(* IEC 61131-3 sources: volt/packages/volt-lsp-iec/test-corpus/awa-palletizer/Device/Plc Logic/Application/Library Manager/L_MC1P_MotionControlBasic, 701 files *)

(* ---- L_MC1P_ABC_STATE.dut ---- *)
TYPE L_MC1P_ABC_STATE :
(
	STANDBY := 0,
	STOP := 1,
	HOMING := 2,
	JOGGING := 3,
	MOVEVEL := 4,
	MOVEABS := 5,
	MOVEREL := 6,
	EXTERNAL := 7,
	ERROR := 8,
	FINISHPOSITIONING := 9
);
END_TYPE

(* ---- L_MC1P_ABORTTRIGGERINPUT.dut ---- *)
TYPE L_MC1P_ABORTTRIGGERINPUT :
STRUCT
	PTRIGGER_REF : POINTER TO MC_TRIGGER_REF;
	EXECUTE : BOOL;
	PAUSEACTIVETP : BOOL;
END_STRUCT
END_TYPE

(* ---- L_MC1P_ABORTTRIGGEROUTPUT.dut ---- *)
TYPE L_MC1P_ABORTTRIGGEROUTPUT :
STRUCT
	DONE : BOOL;
	BUSY : BOOL;
	ERROR : BOOL;
	ERRORID : L_IE1P_Error;
END_STRUCT
END_TYPE

(* ---- L_MC1P_ADDITIONALCONFIGINFO.dut ---- *)
TYPE L_MC1P_ADDITIONALCONFIGINFO :
STRUCT
	LWIDENTDRIVESWITCHOFF : LWORD := 0;
	DWREVISION : DWORD := 0;
	DWMOTORRATEDSPEED : DWORD := 3000;
	LRREFCURRENTMOTOR : LREAL := 0;
	LRREFTORQUEMOTOR : LREAL := 1;
	LRMOTORRATEDTORQUE : LREAL := 1;
	LRTORQUELIMITFACTOR : LREAL := 1;
	LRINERTIAMOTOR : LREAL := 0.01;
	DWMOTORREVOLUTION : DWORD := 1;
	DWENCODERCRC : DWORD := 0;
	XRESETRETAINENCERRORAFTERMAINSWITCH : BOOL;
	XFEEDBACKABSPOSAVAILABLE : BOOL := TRUE;
	XVFCMODE : BOOL := FALSE;
	XTACIA402ADVANCED : BOOL := FALSE;
	WMCTRLMODEDRIVE : USINT := 1;
	XDRIVELOADENCODER : BOOL := FALSE;
	DWDRIVELOADENCODERFEEDBACKCONFIG : DWORD := 0;
	DWDRIVELOADENCODERORIENTATION : DWORD := 0;
	DWDRIVELOADENCODERCRC : DWORD := 0;
	XDEVICETRANSMITTIMESVALID : BOOL;
	LRDEVICETRANSMITTIMEACTPOSMS : LREAL;
	LRDEVICETRANSMITTIMESETPOSMS : LREAL;
END_STRUCT
END_TYPE

(* ---- L_MC1P_ADDITIONALLIMITS.dut ---- *)
TYPE L_MC1P_ADDITIONALLIMITS :
(
	NOTACTIVE := 0,
	ADDITIONALPOSLIMITS := 1
);
END_TYPE

(* ---- L_MC1P_AUTOTUNINGPARA.dut ---- *)
TYPE L_MC1P_AUTOTUNINGPARA :
STRUCT
	MAXVELOCITY : LREAL;
	MAXACCELERATION : LREAL := 0;
	MAXDISTANCE : LREAL := 0;
	MOVEMENTDISTANCE : LREAL := 0;
	STATE : WORD := 0;
	COMMANDIN : USINT;
	VPNFACTOR : WORD;
	TNNFACTOR : WORD;
	VPPFACTOR : WORD;
	VPPFACTOREXT : WORD;
	WAITINGTIME : LREAL;
END_STRUCT
END_TYPE

(* ---- L_MC1P_AVERAGEFILTERSETVALUESINPUT.dut ---- *)
TYPE L_MC1P_AVERAGEFILTERSETVALUESINPUT :
STRUCT
	WFILTERDEPTH : WORD;
	XMANIPULATETORQUE : BOOL := FALSE;
END_STRUCT
END_TYPE

(* ---- L_MC1P_AVERAGEFILTERSETVALUESOUTPUT.dut ---- *)
TYPE L_MC1P_AVERAGEFILTERSETVALUESOUTPUT :
STRUCT
	XINEQOUT : BOOL;
END_STRUCT
END_TYPE

(* ---- L_MC1P_AXIS_STATE.dut ---- *)
TYPE L_MC1P_AXIS_STATE :
(
	ERRORSTOP := 1,
	DISABLED := 2,
	STANDSTILL := 3,
	STOPPING := 4,
	DISCMOTION := 5,
	SYNCMOTION := 6,
	CONTMOTION := 7,
	HOMING := 8,
	SERVICE := 10
);
END_TYPE

(* ---- L_MC1P_AXISBASICCONTROLINPUT_INTERNAL.dut ---- *)
TYPE L_MC1P_AXISBASICCONTROLINPUT_INTERNAL :
STRUCT
	PAXIS : POINTER TO AXIS_REF;
	DISABLEMOVEFUNEXEC : BOOL;
	XDISABLEPOWERCALL : BOOL;
	XREGULATORON : BOOL;
	XRESETERROR : BOOL;
	XENABLEPOSITIVE : BOOL := TRUE;
	XENABLENEGATIVE : BOOL := TRUE;
	XDISABLESWLIMIT : BOOL;
	LROVERRIDE : LREAL := 1.0;
	LROVERRIDEACC : LREAL := 1.0;
	LROVERRIDEJERK : LREAL := 1.0;
	XSTOP : BOOL;
	LRSTOPDEC : LREAL;
	LRSTOPJERK : LREAL;
	XJOGGINGPOS : BOOL;
	XJOGGINGNEG : BOOL;
	LRJOGGINGSETVEL : LREAL := 3600;
	LRJOGGINGSETACC : LREAL := 36000;
	LRJOGGINGSETDEC : LREAL := 36000;
	LRJOGGINGSETJERK : LREAL := 0;
	LRJOGGINGSETJERKDEC : LREAL := 0;
	XCONTINUOUSUPDATE : BOOL;
	XFINISHPOSITIONING : BOOL;
	XQSPAPPLICATION : BOOL;
	XHALT : BOOL;
	XABORT : BOOL;
	XMOVEVELEXECUTE : BOOL;
	XMOVEABSEXECUTE : BOOL;
	XMOVERELEXECUTE : BOOL;
	LRSETPOS_DIST : LREAL;
	LRSETVEL : LREAL := 3600;
	LRSETACC : LREAL := 36000;
	LRSETDEC : LREAL := 36000;
	LRSETJERK : LREAL := 0;
	LRSETJERKDEC : LREAL := 0;
	ESETDIRECTION : MC_DIRECTION := MC_DIRECTION.mcPositiveDirection;
	XHOMEEXECUTE : BOOL;
	LRHOMEPOSITION : LREAL;
	XUSEHOMEEXTPARAMETER : BOOL;
	SCHOMEEXTPARAMETER : L_MC1P_HomeParameter;
	SCHOMEEXTTP : MC_TRIGGER_REF;
	XHOMEABSSWITCH : BOOL;
	XRESETHOMEPOSITION : BOOL;
	XMOVEVELENABLEOFFSETVEL : BOOL;
	LRMOVEVELOFFSETVEL : LREAL;
	XUSEABORTBEHAVIOURFORTM : BOOL;
	LRABORTDEC : LREAL;
	LRABORTJERK : LREAL;
END_STRUCT
END_TYPE

(* ---- L_MC1P_AXISBASICCONTROLINSTANCEDATA.dut ---- *)
TYPE L_MC1P_AXISBASICCONTROLINSTANCEDATA :
STRUCT
	XERROR : BOOL;
	EERRORID : L_IE1P_Error;
	XFUNBUSY : BOOL;
	XFUNDONE : BOOL;
	XFUNCOMMANDABORTED : BOOL;
	EFUNSTATEACT : L_MC1P_ABC_State;
	ABCFUNID : WORD;
	WPOWID : WORD;
	XEXIT : BOOL;
	XMOVEVELEXECUTEOLD : BOOL;
	XMOVEABSEXECUTEOLD : BOOL;
	XMOVERELEXECUTEOLD : BOOL;
	XFINISHPOSITIONINGOLD : BOOL;
	XHOMEEXECUTEOLD : BOOL;
	XJOGGINGNEGOLD : BOOL;
	XJOGGINGPOSOLD : BOOL;
	XSTOPOLD : BOOL;
	XHALTOLD : BOOL;
	XABORTOLD : BOOL;
	XPOWERROROLD : BOOL;
	XDISABLESWLIMITOLD : BOOL;
	XFUNDONEOLD : BOOL;
	XRESETHOMEPOSITIONOLD : BOOL;
	XSAVEMOVEVELDONE : BOOL;
	XACYCLICAXIS : BOOL;
	XQSPAPPLDETECTED : BOOL;
	FBSTOP_EXECUTE : BOOL;
	FBHALT_EXECUTE : BOOL;
	FBABORT_EXECUTE : BOOL;
	FBMOVEABS_EXECUTE : BOOL;
	FBMOVEVEL_EXECUTE : BOOL;
	FBMOVEREL_EXECUTE : BOOL;
	FBFINISHPOSITIONING_XFINISHPOSITIONING : BOOL;
	FBFINISHPOSITIONING_XENABLE : BOOL;
	FBJOG_XJOGPOSITIVE : BOOL;
	FBJOG_XJOGNEGATIVE : BOOL;
	FBHOME_EXECUTE : BOOL;
	FBSTOP_XINUSE : BOOL;
	FBHALT_XINUSE : BOOL;
	FBABORT_XINUSE : BOOL;
	FBMOVEABS_XINUSE : BOOL;
	FBMOVEVEL_XINUSE : BOOL;
	FBMOVEREL_XINUSE : BOOL;
	FBFINISHPOSITIONING_XINUSE : BOOL;
	FBJOG_XINUSE : BOOL;
	FBHOME_XINUSE : BOOL;
	XDRIVEENABLEDOLD_READMOTIONSTATE : BOOL;
	LRACTVELOCITYOLD_READMOTIONSTATE : LREAL;
	LRSETVELOCITYOLD_READMOTIONSTATE : LREAL;
	FBBASEOLD : POINTER TO L_MC1P_Template_ForAxis;
	FBSTOP_FBBASESTATUS : L_MC1P_Template_ForAxis;
	FBHALT_FBBASESTATUS : L_MC1P_Template_ForAxis;
	FBABORT_FBBASESTATUS : L_MC1P_Template_ForAxis;
	FBHOME_FBBASESTATUS : L_MC1P_Template_ForAxis;
	FBJOG_FBBASESTATUS : L_MC1P_Template_ForAxis;
	FBMOVEABS_FBBASESTATUS : L_MC1P_Template_ForAxis;
	FBMOVEVEL_FBBASESTATUS : L_MC1P_Template_ForAxis;
	FBMOVEREL_FBBASESTATUS : L_MC1P_Template_ForAxis;
	FBFINISHPOSITIONING_FBBASESTATUS : L_MC1P_Template_ForAxis;
	FBSETFASTSTOP_FBBASESTATUS : L_MC1P_Template_ForAxis;
	FBSETFASTSTOPINPUT : L_MC1P_SetQuickStopApplInput;
	FBSETFASTSTOP : L_MC1P_SetFastStop_Internal;
	FBSETFASTSTOPOUTPUT : L_MC1P_SetQuickStopApplOutput;
	FBRESET_FBBASESTATUS : L_MC1P_Template_ForAxis;
	FBRESET : L_MC1P_Reset_Internal;
	RESETINPUT : L_MC1P_ResetInput;
	RESETOUTPUT : L_MC1P_ResetOutput;
	FBSETOVERRIDE_FBBASESTATUS : L_MC1P_Template_ForAxis;
	FBSETOVERRIDE : L_MC1P_SetOverride_Internal;
	FBREADMOTIONSTATEINPUT : L_MC1P_ReadMotionStateInput;
	FBREADMOTIONSTATE_FBBASESTATUS : L_MC1P_Template_ForAxis;
	FBREADMOTIONSTATE : L_MC1P_ReadMotionState_Internal;
	FBREADMOTIONSTATEOUTPUT : L_MC1P_ReadMotionStateOutput;
	FBREADAXISERROR_FBBASESTATUS : L_MC1P_Template_ForAxis;
	FBREADAXISERROR : L_MC1P_ReadAxisError_Internal;
	FBREADAXISERRORINPUT : L_MC1P_ReadAxisErrorInput;
	FBREADAXISERROROUTPUT : L_MC1P_ReadAxisErrorOutput;
END_STRUCT
END_TYPE

(* ---- L_MC1P_AXISBASICCONTROLOUTPUT_INTERNAL.dut ---- *)
TYPE L_MC1P_AXISBASICCONTROLOUTPUT_INTERNAL :
STRUCT
	ECONTROLMODE : L_MC1P_ControlMode;
	XISHOMED : BOOL;
	XHWLIMITSWITCHNEG : BOOL;
	XHWLIMITSWITCHPOS : BOOL;
	XSWLIMITENABLED : BOOL;
	XSWLIMITSWITCHNEG : BOOL;
	XSWLIMITSWITCHPOS : BOOL;
	EAXISTYPE : L_MC1P_DriveType;
	EAXISSTATE : L_MC1P_AXIS_STATE := L_MC1P_AXIS_STATE.Disabled;
	XAXISREADY : BOOL;
	XAXISENABLED : BOOL;
	XAXISWARNING : BOOL;
	XAXISERROR : BOOL;
	EAXISERRORID : L_IE1P_Error;
	XDRIVEWARNING : BOOL;
	XDRIVEERROR : BOOL;
	DWDRIVEERRORID : DWORD;
	LRACTPOS : LREAL;
	LRACTVEL : LREAL;
	LRSETPOSOUT : LREAL;
	LRSETVELOUT : LREAL;
	LRACTFOLLOWINGERROR : LREAL;
	XCONSTANTVELOCITY : BOOL;
	XACCELERATING : BOOL;
	XDECELERATING : BOOL;
	XDIRECTIONPOSITIVE : BOOL;
	XDIRECTIONNEGATIVE : BOOL;
	XINPOSITION : BOOL;
	XAXISAVAILABLE : BOOL;
	XSTANDSTILLSETVELOCITY : BOOL;
	XSTANDSTILLACTVELOCITY : BOOL;
	XAXISREADYTOSWITCHON : BOOL;
	XAXISREADYFORMOTION : BOOL;
	XERROR : BOOL;
	EERRORID : L_IE1P_Error;
	XFUNBUSY : BOOL;
	XFUNDONE : BOOL;
	XFUNCOMMANDABORTED : BOOL;
	EFUNSTATEACT : L_MC1P_ABC_State;
	XSTOACTIVE : BOOL;
END_STRUCT
END_TYPE

(* ---- L_MC1P_AXISEXTENSIONTYPES.dut ---- *)
TYPE L_MC1P_AXISEXTENSIONTYPES :
(
	EMPTY := 0,
	HL9400_ECAT := 1,
	HL9400_CAN := 2,
	I500_ECAT := 3,
	I500_CAN := 4,
	I700 := 5,
	I750 := 6,
	I950 := 7,
	I950ADV := 8,
	I950_DRIVE := 9,
	I950_DRIVECIA := 10,
	GENERICDRIVE := 11,
	ENCFREE := 101,
	ENCIO_BPB := 102,
	ENCIO_ECAT := 103,
	ENCI900_ECAT := 104,
	ENCI900_DRIVE := 105,
	ENCI900_DRIVECIA := 106,
	ENCI500_ECAT := 107
);
END_TYPE

(* ---- L_MC1P_AXISFUNCTION.dut ---- *)
TYPE L_MC1P_AXISFUNCTION :
(
	SIMPLEMODE := 1,
	PLI := 2,
	MOL := 3,
	POSCTRLADAPT := 4,
	SPEEDCTRLADAPT := 5,
	SPEEDCTRLLOAD := 6,
	BRAKEGRINDIN := 7,
	BRAKETEST := 8,
	BASICBRAKECTRLONLYINDRIVE := 9,
	FLEXIBLEMAPPING := 10,
	ZEROPULS2NDFEEDBACK := 11,
	FDBSTATUSBITSAVAILABLE := 12,
	AUTOTUNING := 13,
	PARSAVEINDRIVE := 14,
	WAITFORAXISDETECTION := 15
);
END_TYPE

(* ---- L_MC1P_AXISGUID.dut ---- *)
TYPE L_MC1P_AXISGUID :
STRUCT
	ADWDATA : ARRAY [1..4] OF DWORD;
END_STRUCT
END_TYPE

(* ---- L_MC1P_AXISINTERFACEINPUT.dut ---- *)
TYPE L_MC1P_AXISINTERFACEINPUT :
STRUCT
	XENABLE : BOOL;
	EXTCONTROLLER : L_MC1P_IControllerInterface;
END_STRUCT
END_TYPE

(* ---- L_MC1P_AXISINTERFACEOUTPUT.dut ---- *)
TYPE L_MC1P_AXISINTERFACEOUTPUT :
STRUCT
	XVALID : BOOL;
	XBUSY : BOOL;
	XERROR : BOOL;
	EERRORID : L_IE1P_Error;
END_STRUCT
END_TYPE

(* ---- L_MC1P_AXISPROPERTIES.dut ---- *)
TYPE L_MC1P_AXISPROPERTIES :
STRUCT
	XVIRTUAL : BOOL := FALSE;
	XTPSUPPORTED : BOOL := FALSE;
	XTPWITHTIMESTAMP : BOOL := FALSE;
	SNTPMAXCHANNEL : SINT := 0;
	XSUPPORTBRAKE : BOOL := FALSE;
	XSUPPORTDCBRAKE : BOOL := FALSE;
	XCHECKCOMMUNICATIONSTATE : BOOL := TRUE;
	XDRIVEHOMINGSUPPORTED : BOOL := FALSE;
	XTACIAADVANCED : BOOL := FALSE;
	BYDELAYLIMITDRIVEOPERATIONENABLED : BYTE := 2;
	LRTRANSMITCYCLESACTPOS : LREAL;
	LRTRANSMITCYCLESSETPOS : LREAL;
	DWTPDELAYACTPOS : DWORD;
	XFORWARDECATSLAVEERROR : BOOL := FALSE;
	XFORCEACYCLICMODE : BOOL := FALSE;
	WOFFSETDRIVEPARA : WORD := 0;
END_STRUCT
END_TYPE

(* ---- L_MC1P_AXISRETAININFO.dut ---- *)
TYPE L_MC1P_AXISRETAININFO :
STRUCT
	MEMTYPE : BYTE;
	MEMVERSION : BYTE;
	MEMLENGTH : WORD;
END_STRUCT
END_TYPE

(* ---- L_MC1P_AXISRETAININFORMATION.dut ---- *)
TYPE L_MC1P_AXISRETAININFORMATION :
STRUCT
	AXISGUID : L_MC1P_AxisGUID;
	ITFRETAIN : L_MC1P_IRetainFunction;
	PDATA : POINTER TO DWORD;
	PDATAMIRROR : POINTER TO DWORD;
END_STRUCT
END_TYPE

(* ---- L_MC1P_AXISSIMIODATA.dut ---- *)
TYPE L_MC1P_AXISSIMIODATA :
STRUCT
	XSTO : BOOL;
	XDIGIN1 : BOOL;
	XDIGIN2 : BOOL;
	XSTIMULATEERROR : BOOL;
	DWERRORCODE : DWORD;
	XQSPONERROR : BOOL;
	XSTIMULATEWARNING : BOOL;
	DWWARNINGCODE : DWORD;
	ETPMODE : UINT := 0;
	LRTPDISTANCE : LREAL;
	LRTPDISTANCEINTERNAL : LREAL;
	XSTIMULATEFEEDBACKCHANGED : BOOL;
END_STRUCT
END_TYPE

(* ---- L_MC1P_AXISSIMULATIONPDODATAFROMDRIVE.dut ---- *)
TYPE L_MC1P_AXISSIMULATIONPDODATAFROMDRIVE :
STRUCT
	UICIASTATUSWORD : UINT;
	UILENZESTATUSWORD : UINT;
	SIMODEOFOPERATIONDISP : SINT;
	UIERRORCODE : UINT;
	UITEXTREFID : UINT;
	DIVELACTVALUE : DINT;
	ITORQUEACTVALUE : INT;
	DIPOSACTVALUE : DINT;
	DIFOLLOWINGERRORACTVALUE : DINT;
	IVLACTUALVEL : INT;
	UITPSTATUS : UINT;
	DITPPOS1POSVALUE : DINT;
	DITPPOS1NEGVALUE : DINT;
	DITPPOS2POSVALUE : DINT;
	DITPPOS2NEGVALUE : DINT;
	UILENZESTATUSWORD2 : UINT;
	UDIDIGITALINPUTS : UDINT;
END_STRUCT
END_TYPE

(* ---- L_MC1P_AXISSIMULATIONPDODATAFROMDRIVESCALED.dut ---- *)
TYPE L_MC1P_AXISSIMULATIONPDODATAFROMDRIVESCALED :
STRUCT
	UICIASTATUSWORD : UINT;
	UILENZESTATUSWORD : UINT;
	SIMODEOFOPERATIONDISP : SINT;
	UIERRORCODE : UINT;
	UITEXTREFID : UINT;
	LRVELACTVALUE : LREAL;
	LRTORQUEACTVALUE : LREAL;
	LRPOSACTVALUE : LREAL;
	LRFOLLOWINGERRORACTVALUE : LREAL;
	UITPSTATUS : UINT;
	LRTPPOS1POSVALUE : LREAL;
	LRTPPOS1NEGVALUE : LREAL;
	LRTPPOS2POSVALUE : LREAL;
	LRTPPOS2NEGVALUE : LREAL;
	UILENZESTATUSWORD2 : UINT;
	UDIDIGITALINPUTS : UDINT;
END_STRUCT
END_TYPE

(* ---- L_MC1P_AXISSIMULATIONPDODATATODRIVE.dut ---- *)
TYPE L_MC1P_AXISSIMULATIONPDODATATODRIVE :
STRUCT
	UICTRLWORD : UINT;
	UILENZECTRLWORD : UINT;
	SIMODEOFOPERATION : SINT;
	ITORQUEOFFSET : INT;
	DITARGETPOSITION : DINT;
	DIVELOCITYOFFSET : DINT;
	ISPDCTRL_ILOADVALUE : INT;
	ITARGETTORQUE : INT;
	DITARGETVELOCITY : DINT;
	IVLTARGETVEL : INT;
	UITPFUNCTION1 : UINT;
	UIPOSTORQUELIMIT : UINT;
	UINEGTORQUELIMIT : UINT;
	DIUPPERSPEEDLIMIT : DINT;
	DILOWERSPEEDLIMIT : DINT;
END_STRUCT
END_TYPE

(* ---- L_MC1P_AXISSIMULATIONPDODATATODRIVESCALED.dut ---- *)
TYPE L_MC1P_AXISSIMULATIONPDODATATODRIVESCALED :
STRUCT
	UICTRLWORD : UINT;
	UILENZECTRLWORD : UINT;
	SIMODEOFOPERATION : SINT;
	LRSETPOSITION : LREAL;
	LRSETVELOCITY : LREAL;
	LRSETTORQUE : LREAL;
	LRSPDCTRL_ILOADVALUE : LREAL;
	LRVLTARGETVELOCITY : LREAL;
	UITPFUNCTION1 : UINT;
	LRPOSTORQUELIMIT : LREAL;
	LRNEGTORQUELIMIT : LREAL;
	LRUPPERSPEEDLIMIT : LREAL;
	LRLOWERSPEEDLIMIT : LREAL;
END_STRUCT
END_TYPE

(* ---- L_MC1P_AXISSIMULATIONSDODATA.dut ---- *)
TYPE L_MC1P_AXISSIMULATIONSDODATA :
STRUCT
	LRRATEDMOTORTORQUE : LREAL := 0.6;
	LRRATEDMOTORSPEED : LREAL := 4050;
	LRINERTIAMOTOR : LREAL := 0.14;
	LRINERTIALOAD : LREAL := 0;
	LRMOTORRATEDCURRENT : LREAL := 1.8;
	LRMAXMOTORSPEED : LREAL := 6075;
	BYMCTRLMODE : BYTE := 1;
	LRVP_SPEEDCTRL : LREAL := 0.00045;
	LRTN_SPEEDCTRL : LREAL := 12.8;
	LRVP_POSCTRL : LREAL := 28.4;
	LRPOSCTRLOUTPUTLIMITATION : LREAL := 480000;
	UIINSABILITYVALUE : UINT;
	UIINSABILITYINDICATOR : USINT;
	USISWITCHINGFREQUENCY : USINT := 1;
	LRPOSCTRLADAPT : LREAL := 100.0;
	LRSPEEDCTRLADAPT : LREAL := 100.0;
	LRMAXTORQUE : LREAL := 250.0;
	LRSPEEDFILTERTIME : LREAL := 0.3;
	WNBRORREVOLUTION : WORD := 1;
	DWINKPERREV : DWORD := 65536;
	DWENCODERCRC : DWORD := 1234;
	DWENCODERCRCLOAD : DWORD := 4567;
	USIBRAKEMODE : USINT := 2;
	UIBRAKESRCOFSTARTINGTORQUE : UINT := 1;
	LRBRAKEDETECTEDSTARTINGTORQUE : LREAL := 0;
	LRBRAKERELEASINGTIME : LREAL := 0.1;
	LRBRAKECLOSINGTIME : LREAL := 0.1;
	USIBRAKEOVERRIDE : USINT := 0;
	LRSTARTTORQUE : LREAL;
	UIBRAKELOGICSTATE : UINT;
	UICONTROLMODECIA402ADVANCED : UINT := 0;
	LRVP_LOADPOSCTRL : LREAL := 20.0;
	SIIPOTIMEEXP : SINT;
	USIIPOTIME : USINT;
	UIQSPOPTION : UINT;
	UDIPOSITIONREACHEDWINDOW : UDINT := 1000;
	UDIQSPDECELERATION : UDINT := 2147483647;
	DWREVISIONNBR : DWORD := 16#20000;
	DWFIRSTSYNCTIME : DWORD;
	USISPEEDERRORRESPONSE : USINT;
	SSWVERSION : STRING(50) := '1.7.5.2420 (release)';
	USIDISABLEPDOS : USINT;
	USIDRIVECOMMAND_0X2825 : USINT;
	UDIMAINSWITCHINGCYCLES_0X2D81_4 : UDINT := 666;
	USIPOSSETMODE_0X2984 : USINT;
	LRVLACCDELTASPEED : LREAL := 0;
	LRVLACCDELTATIME : LREAL := 10;
	LRVLDECDELTASPEED : LREAL := 0;
	LRVLDECDELTATIME : LREAL := 0;
	BYDISABLEDEVICE : BYTE;
	DIADDSPEEDLIMITATION : DINT := 0;
	AUIGAINCHARACTERISTIC : ARRAY [1..11] OF WORD := [10, 100, 100, 100, 1000, 100, 2000, 100, 5000, 100, 0];
END_STRUCT
END_TYPE

(* ---- L_MC1P_AXISSLOT.dut ---- *)
TYPE L_MC1P_AXISSLOT :
(
	AXISA := 16#0,
	AXISB := 16#800
);
END_TYPE

(* ---- L_MC1P_AXISTYPE.dut ---- *)
TYPE L_MC1P_AXISTYPE :
(
	UNKNOWN := 0,
	AXISREF := 1,
	AXISKINEMATIC := 2,
	AXISGROUP := 3
);
END_TYPE

(* ---- L_MC1P_BACKLASHCONTACTSTATE.dut ---- *)
TYPE L_MC1P_BACKLASHCONTACTSTATE :
(
	NOCONTACT := 0,
	NEGATIVECONTACT := 1,
	POSITIVECONTACT := 2
);
END_TYPE

(* ---- L_MC1P_BASICACTUATINGSPEEDINPUT.dut ---- *)
TYPE L_MC1P_BASICACTUATINGSPEEDINPUT :
STRUCT
	XENABLEINTERNALCONTROL : BOOL := FALSE;
	XREGULATORON : BOOL := FALSE;
	XRESETERROR : BOOL := FALSE;
	XSETDRIVEQSP : BOOL := FALSE;
	XENABLESETVEL : BOOL := FALSE;
	XINVERTDIRECTION : BOOL := FALSE;
	LRSETVEL : LREAL := 0.0;
	LRSETACC : LREAL := 0.0;
	LRSETDEC : LREAL := 0.0;
END_STRUCT
END_TYPE

(* ---- L_MC1P_BASICACTUATINGSPEEDOUTPUT.dut ---- *)
TYPE L_MC1P_BASICACTUATINGSPEEDOUTPUT :
STRUCT
	XINTERNALCONTROLACTIVE : BOOL;
	XBUSY : BOOL;
	XERROR : BOOL;
	EERRORID : L_IE1P_Error;
	XCOMMUNICATIONOK : BOOL;
	XAXISREADY : BOOL;
	XAXISENABLED : BOOL;
	XDRIVEWARNING : BOOL;
	XDRIVEERROR : BOOL;
	DWDRIVEERRORID : DWORD;
	XDRIVEQSPACTIVE : BOOL;
	LRACTVEL : LREAL;
	XDIRECTIONPOSITIVE : BOOL;
	XDIRECTIONNEGATIVE : BOOL;
	WDIGITALINPUTS : WORD;
END_STRUCT
END_TYPE

(* ---- L_MC1P_BRAKEAUTOSTATE.dut ---- *)
TYPE L_MC1P_BRAKEAUTOSTATE :
(
	AS_IDLE,
	AS_RAMPDOWN,
	AS_CLOSINGBRAKE,
	AS_INITBRAKECLOSE,
	AS_BRAKECLOSED,
	AS_RELEASINGBRAKE,
	AS_SUPERVISORMODE,
	AS_DIRECTCONTROL
);
END_TYPE

(* ---- L_MC1P_BRAKECMDBRAKEGRINDINPARA.dut ---- *)
TYPE L_MC1P_BRAKECMDBRAKEGRINDINPARA :
STRUCT
	MOTORSPEED : INT := 1000;
	RAMPTIME : INT := 1000;
	ONTIME : INT := 500;
	OFFTIME : INT := 500;
	CYCLES : WORD := 4;
	GRINDINCONTROL : BYTE;
	MODE : USINT;
	CYCLESOUT : WORD;
	STATE : WORD;
	POSLIMIT1 : LREAL;
	POSLIMIT2 : LREAL;
END_STRUCT
END_TYPE

(* ---- L_MC1P_BRAKECMDBRAKETESTPARA.dut ---- *)
TYPE L_MC1P_BRAKECMDBRAKETESTPARA :
STRUCT
	MOTORTORQUE : DINT := 0;
	RAMPTIME : INT := 1000;
	HOLDTIME : INT := 4000;
	POSTHRESHOLD : INT;
	STATE : WORD := 0;
	WBRAKETESTMODE : USINT;
END_STRUCT
END_TYPE

(* ---- L_MC1P_BRAKECTRL.dut ---- *)
TYPE L_MC1P_BRAKECTRL :
STRUCT
	XDISABLEPHIERR : BOOL;
	XBRAKEFQSP : BOOL;
	XTORQUETIMEOUT : BOOL;
	XRELEASED : BOOL;
	XOUTPUTRELEASEOLD : BOOL;
	XOBSERVE : BOOL;
	XMODULENOTOK : BOOL;
	XEXTSIGNOTOK : BOOL;
	XMODULEFEEDBACK : BOOL;
	XBRAKEOPENED : BOOL;
	XBRAKECLOSED : BOOL;
	XINVERTBRAKE : BOOL;
	XINVERTBRAKEOLD : BOOL;
	XUVDETECTEDOLD : BOOL;
	XACTSPEEDBELOWMINSPEED : BOOL;
	XBIT15 : BOOL;
END_STRUCT
END_TYPE

(* ---- L_MC1P_BRAKEERRORCODES.dut ---- *)
TYPE L_MC1P_BRAKEERRORCODES :
(
	EC_POSITIONDRIFT := 3,
	EC_POSITIONDRIFTCINH := 11,
	EC_RAMPWATCH := 4,
	EC_ERRORMODULE := 5,
	EC_ERROREXTSIGNAL := 13,
	EC_ERRORTORQUETIMEOUT := 18,
	EC_ERRORBRAKESTATEINVALID := 19,
	EC_ERRORBRAKEMODEINVALID := 20,
	EC_TORQUELIMITED := 30
);
END_TYPE

(* ---- L_MC1P_BRAKEGRINDININPUT.dut ---- *)
TYPE L_MC1P_BRAKEGRINDININPUT :
STRUCT
	XEXECUTE : BOOL;
	EMODE : L_MC1P_GrindInMode := L_MC1P_GrindInMode.CwCcw;
	EADDITIONALLIMITS : L_MC1P_AdditionalLimits := L_MC1P_AdditionalLimits.NotActive;
	LRPOSLIMIT1 : LREAL := 0;
	LRPOSLIMIT2 : LREAL := 0;
	LRMOTORSPEED : LREAL := 60.0;
	LRRAMPTIME : LREAL := 1.0;
	LRONTIME : LREAL := 0.5;
	LROFFTIME : LREAL := 0.5;
	WCYCLES : WORD := 4;
	XEXTERNALFAN : BOOL := FALSE;
	XFINISHINSTARTPOS : BOOL := FALSE;
	XUSEAXISPARAMETER : BOOL := FALSE;
	XDISABLEHOMEPOSCHECK : BOOL;
	XGRINDINVELOCITYMODE : BOOL;
	XCYCLESSETBYPARAMETER : BOOL;
	WCYCLESCW : WORD := 2;
	WCYCLESCCW : WORD := 2;
	XALLOWEXECUTIONFORKINEMATICSLAVE : BOOL;
	XABORT : BOOL;
END_STRUCT
END_TYPE

(* ---- L_MC1P_BRAKEGRINDINOUTPUT.dut ---- *)
TYPE L_MC1P_BRAKEGRINDINOUTPUT :
STRUCT
	XDONE : BOOL;
	XBUSY : BOOL;
	XACTIVE : BOOL;
	XCOMMANDABORTED : BOOL;
	XERROR : BOOL;
	EERRORID : L_IE1P_Error;
	WCYCLESOUT : WORD;
	ESTATE : L_MC1P_BrakeGrindInState := L_MC1P_BrakeGrindInState.NotActive;
	XGRINDINABORTEDINSTANDSTILL : BOOL;
END_STRUCT
END_TYPE

(* ---- L_MC1P_BRAKEGRINDINSTATE.dut ---- *)
TYPE L_MC1P_BRAKEGRINDINSTATE :
(
	NOTACTIVE := 0,
	INIT := 1,
	BRAKEGRINDIN := 3,
	DONE := 4,
	ERROR := 5,
	ABORTED := 6,
	BRAKEGRINDINFOLLOWER := 20
);
END_TYPE

(* ---- L_MC1P_BRAKEINTERFACEINPUT.dut ---- *)
TYPE L_MC1P_BRAKEINTERFACEINPUT :
STRUCT
	XENABLE : BOOL;
	XRELEASEBRAKE : BOOL;
	LRTORQUEADD : LREAL;
	XBRAKEMODEACTIVATE : BOOL;
	EBRAKEMODE : L_MC1P_BrakeMode;
END_STRUCT
END_TYPE

(* ---- L_MC1P_BRAKEINTERFACEOUTPUT.dut ---- *)
TYPE L_MC1P_BRAKEINTERFACEOUTPUT :
STRUCT
	XVALID : BOOL;
	XBUSY : BOOL;
	XERROR : BOOL;
	EERRORID : L_IE1P_Error;
	XBRAKERELEASEOUT : BOOL;
	XBRAKERELEASED : BOOL;
	LRACTTORQUE : LREAL;
	LRSTARTINGTORQUESAVED : LREAL;
	LRSTARTINGTORQUEEFFECTIVE : LREAL;
	EBRAKEMODEACTIVE : L_MC1P_BrakeMode;
END_STRUCT
END_TYPE

(* ---- L_MC1P_BRAKELOGICSTATE.dut ---- *)
TYPE L_MC1P_BRAKELOGICSTATE :
(
	OFF := 0,
	WAITON := 1,
	SELECTPRETORQUE := 10,
	LOADPRETORQUE := 11,
	OPENBRAKE := 20,
	OPERATION := 30,
	CLOSEBRAKE := 40,
	TURNOFF := 50
);
END_TYPE

(* ---- L_MC1P_BRAKEMODE.dut ---- *)
TYPE L_MC1P_BRAKEMODE :
(
	OFF := 0,
	MANUALCONTROL_PLC := 1,
	AUTOMATIC_PLC := 2
);
END_TYPE

(* ---- L_MC1P_BRAKEOUTSTATE.dut ---- *)
TYPE L_MC1P_BRAKEOUTSTATE :
STRUCT
	XBRAKECONTROLACTIVE : BOOL;
	XMODULEOPERATION : BOOL;
	XBRAKEOUTSTATE : BOOL;
	XTORQUECTRLACTIVE : BOOL;
	XBRAKECINH : BOOL;
	XERRORACTIVE : BOOL;
	XGRINDINACTIVE : BOOL;
	XTORQUETESTACTIVE : BOOL;
	XMANOPERATION : BOOL;
	XAUTOPERATION : BOOL;
	XERROREXTFEEDBACK : BOOL;
	XERRORPOSDRIFT : BOOL;
	XERRORBRAKEMODULE : BOOL;
	XINFOTIMEOUTACTIVATE : BOOL;
	XGRINDINDONE : BOOL;
	XTORQUETESTDONE : BOOL;
	XERRORTORQUECTRL : BOOL;
	XACTSPEEDBELOWMIN : BOOL;
	XERRORTORQUELIMITED : BOOL;
END_STRUCT
END_TYPE

(* ---- L_MC1P_BRAKEPARA.dut ---- *)
TYPE L_MC1P_BRAKEPARA :
STRUCT
	LRRELEASETIME : LREAL;
	LRACTIVATIONTIME : LREAL;
	DWBRAKEMODE : DWORD;
	ESELBRAKEMODE : DWORD;
	LRSAMPLEDBRAKETORQUE : LREAL;
	LREFFECTIVESTARTINGTORQUE : LREAL;
	ALRMSTARTVALUE : ARRAY [1..2] OF LREAL;
	LRBRAKERAMPTIME : LREAL;
	XBRAKEACCDEPENDING : BOOL;
	WSOURCESTARTVALUE : WORD;
END_STRUCT
END_TYPE

(* ---- L_MC1P_BRAKESTATE.dut ---- *)
TYPE L_MC1P_BRAKESTATE :
(
	EBS_DEFAULT := 0,
	EBS_BRAKECLOSED,
	EBS_BRAKEOPEN,
	EBS_BRAKESWITCHING,
	EBS_BRAKEOBSERVATION,
	EBS_BRAKEAUTO,
	EBS_BRAKEAUTOGSB,
	EBS_BRAKEAUTOSUPERVISOR,
	EBS_BRAKEMANUAL,
	EBS_BRAKEOFF,
	EBS_STATESWITCH,
	EBS_STATEOPERATION
);
END_TYPE

(* ---- L_MC1P_BRAKETESTINPUT.dut ---- *)
TYPE L_MC1P_BRAKETESTINPUT :
STRUCT
	XEXECUTE : BOOL;
	LRMOTORTORQUE : LREAL := 0;
	LRRAMPTIME : LREAL := 1.0;
	LRHOLDTIME : LREAL := 4.0;
	LRPOSTHRESHOLD : LREAL;
	EDIRECTION : MC_DIRECTION := MC_DIRECTION.mcCurrentDirection;
	EMODE : L_MC1P_BrakeTestMode := L_MC1P_BrakeTestMode.NoLoadTorque;
	XUSEAXISPARAMETER : BOOL := FALSE;
	XABORT : BOOL;
	XALLOWEXECUTIONFORKINEMATICSLAVE : BOOL;
END_STRUCT
END_TYPE

(* ---- L_MC1P_BRAKETESTMODE.dut ---- *)
TYPE L_MC1P_BRAKETESTMODE :
(
	NOLOADTORQUE := 0,
	LOADTORQUEIDENTIFICATION := 1
);
END_TYPE

(* ---- L_MC1P_BRAKETESTOUTPUT.dut ---- *)
TYPE L_MC1P_BRAKETESTOUTPUT :
STRUCT
	XDONE : BOOL;
	XBUSY : BOOL;
	XACTIVE : BOOL;
	XCOMMANDABORTED : BOOL;
	XERROR : BOOL;
	EERRORID : L_IE1P_Error;
	LRIDENTIFIEDTORQUE : LREAL;
	LRACTPOSTHRESHOLD : LREAL;
	LRACTMOTORTORQUE : LREAL;
	ESTATE : L_MC1P_BrakeTestState := L_MC1P_BrakeTestState.NotActive;
END_STRUCT
END_TYPE

(* ---- L_MC1P_BRAKETESTSTATE.dut ---- *)
TYPE L_MC1P_BRAKETESTSTATE :
(
	NOTACTIVE := 0,
	INIT := 1,
	TORQUEIDENTIFICATION := 2,
	BRAKETEST := 3,
	DONE := 4,
	ERROR := 5,
	ABORTED := 6,
	BRAKETESTFOLLOWER := 20
);
END_TYPE

(* ---- L_MC1P_BUFFERDATA.dut ---- *)
TYPE L_MC1P_BUFFERDATA :
STRUCT
	LRBUFFERPOSITIONPOS : LREAL;
	LRBUFFERPOSITIONNEG : LREAL;
	LRBUFFERVELPOS : LREAL;
	LRBUFFERVELNEG : LREAL;
END_STRUCT
END_TYPE

(* ---- L_MC1P_CHANGEMACHINEDATAINPUT.dut ---- *)
TYPE L_MC1P_CHANGEMACHINEDATAINPUT :
STRUCT
	XEXECUTE : BOOL;
	XSETFEEDCONSTANT : BOOL;
	LRFEEDCONSTANT : LREAL := 360.0;
	XSETGEARFACTOR : BOOL;
	DWGEARDENOMINATOR : DWORD := 1;
	DWGEARNUMERATOR : DWORD := 1;
	XSETADDGEARFACTOR : BOOL;
	DWADDGEARDENOMINATOR : DWORD := 1;
	DWADDGEARNUMERATOR : DWORD := 1;
	XSETPOSRESOLUTION : BOOL;
	DWPOSRESOLUTION : DWORD := 65536;
	XSETORIENTATION : BOOL;
	XORIENTATION : BOOL := FALSE;
	XSETTRAVERSINGRANGE : BOOL;
	ETRAVERSINGRANGE : L_MC1P_TraversingRange := L_MC1P_TraversingRange.Limited;
	XSETCYCLELENGTH : BOOL;
	LRCYCLELENGTH : LREAL := 360.0;
END_STRUCT
END_TYPE

(* ---- L_MC1P_CHANGEMACHINEDATAOUTPUT.dut ---- *)
TYPE L_MC1P_CHANGEMACHINEDATAOUTPUT :
STRUCT
	XDONE : BOOL;
	XBUSY : BOOL;
	XERROR : BOOL;
	EERRORID : L_IE1P_Error;
END_STRUCT
END_TYPE

(* ---- L_MC1P_CINHHANDLINGINPUT.dut ---- *)
TYPE L_MC1P_CINHHANDLINGINPUT :
STRUCT
	XENABLE : BOOL;
	XSTAYINLASTSTATE : BOOL;
	XMOVELASTSETPOS : BOOL;
	LRWINDOWPOS : LREAL;
	LRWINDOWNEG : LREAL;
	LRSETVEL : LREAL;
	LRSETACC : LREAL;
	LRSETDEC : LREAL;
	LRSETJERK : LREAL;
	EDIRECTION : MC_DIRECTION;
END_STRUCT
END_TYPE

(* ---- L_MC1P_CINHHANDLINGOUTPUT.dut ---- *)
TYPE L_MC1P_CINHHANDLINGOUTPUT :
STRUCT
	XDONE : BOOL;
	XBUSY : BOOL;
	XACTIVE : BOOL;
	XERROR : BOOL;
	EERRORID : L_IE1P_Error;
	XREADYTOCONTINUE : BOOL;
	XINSIDEPOSWINDOW : BOOL;
	XINSIDEACTPOSWINDOW : BOOL;
	EAXISSTATEREAL : L_MC1P_AXIS_STATE := L_MC1P_AXIS_STATE.Disabled;
	LRDISTANCE : LREAL;
END_STRUCT
END_TYPE

(* ---- L_MC1P_CLASSID.dut ---- *)
TYPE L_MC1P_CLASSID :
(
	AXIS_REF := (L_MC1P_Internal.cdiEnumStartValue + 2),
	AXISBASICCONTROLV2 := (L_MC1P_Internal.cdiEnumStartValue + 3)
);
END_TYPE

(* ---- L_MC1P_COMPENSATIONMODE.dut ---- *)
TYPE L_MC1P_COMPENSATIONMODE :
(
	OFF := 0,
	AUTOMATICSET := 1,
	AUTOMATICACT := 2,
	MANUALLY := 3
);
END_TYPE

(* ---- L_MC1P_CONTROLAXIS.dut ---- *)
TYPE L_MC1P_CONTROLAXIS :
STRUCT
	XENABLEOPERATION : BOOL;
	XRESETERROR : BOOL;
	XQSPAPPLICATION : BOOL;
	XJOGPOS : BOOL;
	XJOGNEG : BOOL;
	LRJOGOVERRIDE : LREAL := 1.0;
	LRJOGDISTANCE : LREAL := 10;
	XRESETHOMEPOSITION : BOOL;
END_STRUCT
END_TYPE

(* ---- L_MC1P_CONTROLMODE.dut ---- *)
TYPE L_MC1P_CONTROLMODE :
(
	POSCTRLDRIVE := 0,
	POSCTRLPLC := 1,
	SPEEDCTRLDRIVE := 10,
	TORQUECTRLDRIVE := 20
);
END_TYPE

(* ---- L_MC1P_CONTROLMODESET.dut ---- *)
TYPE L_MC1P_CONTROLMODESET :
(
	POSCTRLDRIVE := 0,
	POSCTRLPLC := 1,
	SPEEDCTRLDRIVE := 10
);
END_TYPE

(* ---- L_MC1P_CTRLABC.dut ---- *)
TYPE L_MC1P_CTRLABC :
STRUCT
	XREGULATORON : BOOL;
	XRESETERROR : BOOL;
	XENABLEPOSITIVE : BOOL := TRUE;
	XENABLENEGATIVE : BOOL := TRUE;
	XDISABLESWLIMIT : BOOL;
	LROVERRIDE : LREAL := 1.0;
	LROVERRIDEACC : LREAL := 1.0;
	LROVERRIDEJERK : LREAL := 1.0;
	XSTOP : BOOL;
	LRSTOPDEC : LREAL := 360000;
	LRSTOPJERK : LREAL := 0;
	XJOGGINGPOS : BOOL;
	XJOGGINGNEG : BOOL;
	XCONTINUOUSUPDATE : BOOL;
	XMOVEVELEXECUTE : BOOL;
	XMOVEABSEXECUTE : BOOL;
	XMOVERELEXECUTE : BOOL;
	XHALT : BOOL;
	LRSETPOS_DIST : LREAL;
	ESETDIRECTION : MC_DIRECTION := MC_DIRECTION.mcPositiveDirection;
	XHOMEEXECUTE : BOOL;
	LRHOMEPOSITION : LREAL;
	XUSEHOMEEXTPARAMETER : BOOL;
	SCHOMEEXTPARAMETER : L_MC1P_HomeParameter;
	SCHOMEEXTTP : MC_TRIGGER_REF;
	XHOMEABSSWITCH : BOOL;
END_STRUCT
END_TYPE

(* ---- L_MC1P_CYCLICPARAMETERACCESSREADINPUT.dut ---- *)
TYPE L_MC1P_CYCLICPARAMETERACCESSREADINPUT :
STRUCT
	XENABLE : BOOL;
	WINDEX : WORD;
	USISUBINDEX : USINT;
	USISIZE : USINT;
	XSIGNED : BOOL := FALSE;
	LRSCALEFACTOR : LREAL := 1;
END_STRUCT
END_TYPE

(* ---- L_MC1P_CYCLICPARAMETERACCESSREADOUTPUT.dut ---- *)
TYPE L_MC1P_CYCLICPARAMETERACCESSREADOUTPUT :
STRUCT
	XVALID : BOOL;
	XBUSY : BOOL;
	XERROR : BOOL;
	EERRORID : L_IE1P_Error;
	LRDATA : LREAL;
END_STRUCT
END_TYPE

(* ---- L_MC1P_CYCLICPARAMETERACCESSWRITEINPUT.dut ---- *)
TYPE L_MC1P_CYCLICPARAMETERACCESSWRITEINPUT :
STRUCT
	XENABLE : BOOL;
	WINDEX : WORD;
	USISUBINDEX : USINT;
	USISIZE : USINT;
	XSIGNED : BOOL := FALSE;
	LRSCALEFACTOR : LREAL := 1;
	LRDATA : LREAL;
END_STRUCT
END_TYPE

(* ---- L_MC1P_CYCLICPARAMETERACCESSWRITEOUTPUT.dut ---- *)
TYPE L_MC1P_CYCLICPARAMETERACCESSWRITEOUTPUT :
STRUCT
	XVALID : BOOL;
	XBUSY : BOOL;
	XERROR : BOOL;
	EERRORID : L_IE1P_Error;
END_STRUCT
END_TYPE

(* ---- L_MC1P_DELAYSETVALUESINPUT.dut ---- *)
TYPE L_MC1P_DELAYSETVALUESINPUT :
STRUCT
	LRDELAYTIME : LREAL := 0.1;
	XEXECUTIONINDEXINTERN : BOOL;
END_STRUCT
END_TYPE

(* ---- L_MC1P_DELAYSETVALUESOUTPUT.dut ---- *)
TYPE L_MC1P_DELAYSETVALUESOUTPUT :
STRUCT
	XINEQOUT : BOOL;
END_STRUCT
END_TYPE

(* ---- L_MC1P_DEVICECLASS.dut ---- *)
TYPE L_MC1P_DEVICECLASS :
(
	VIRTUALAXIS := 0,
	REALAXIS := 1,
	ENCODERAXIS := 2
);
END_TYPE

(* ---- L_MC1P_DIRECTION.dut ---- *)
TYPE L_MC1P_DIRECTION :
(
	BOTH := 0,
	DIRECTIONMASTER := 1
);
END_TYPE

(* ---- L_MC1P_DISABLESWLIMITINPUT.dut ---- *)
TYPE L_MC1P_DISABLESWLIMITINPUT :
STRUCT
	XENABLE : BOOL;
END_STRUCT
END_TYPE

(* ---- L_MC1P_DISABLESWLIMITOUTPUT.dut ---- *)
TYPE L_MC1P_DISABLESWLIMITOUTPUT :
STRUCT
	XBUSY : BOOL;
	XERROR : BOOL;
	EERRORID : L_IE1P_Error;
END_STRUCT
END_TYPE

(* ---- L_MC1P_DRIVESPECIFICCONTAINER.dut ---- *)
TYPE L_MC1P_DRIVESPECIFICCONTAINER :
UNION
	PDATA : POINTER TO BYTE;
	BASIC : POINTER TO L_MC1P_DriveSpecific_Basic;
	CIA402 : POINTER TO L_MC1P_DriveSpecific_CiA402;
	I500 : POINTER TO L_MC1P_DriveSpecific_i500;
	I700 : POINTER TO L_MC1P_DriveSpecific_i700;
	I750 : POINTER TO L_MC1P_DriveSpecific_i750;
	I950 : POINTER TO L_MC1P_DriveSpecific_i950;
	I950ADV : POINTER TO L_MC1P_DriveSpecific_i950Adv;
	I950DRIVE : POINTER TO L_MC1P_DriveSpecific_i950_Drive;
	HL9400 : POINTER TO L_MC1P_DriveSpecific_9400HL;
	ENC : POINTER TO L_MC1P_DriveSpecific_Enc;
	ENC_BPB : POINTER TO L_MC1P_DriveSpecific_Enc_Bpb;
	ENC_FREE : POINTER TO L_MC1P_DriveSpecific_Enc_Free;
	ENC_I950 : POINTER TO L_MC1P_DriveSpecific_Enc_i950;
	ENC_I500 : POINTER TO L_MC1P_DriveSpecific_Enc_i500;
	ENC_IOECAT : POINTER TO L_MC1P_DriveSpecific_Enc_IOETC;
END_UNION
END_TYPE

(* ---- L_MC1P_DRIVESTATECOLLECTION.dut ---- *)
TYPE L_MC1P_DRIVESTATECOLLECTION :
STRUCT
	BYDRIVESTATE : BYTE;
	XDRIVETESTMODEACTIVE : BOOL;
	XDRIVEQSPACTIVE : BOOL;
	XDRIVEQSPDONE : BOOL;
	XSTOACTIVE : BOOL;
	XCINHACTIVE : BOOL;
	XVOLTAGEENABLED : BOOL;
	XUSEQSPDRIVEINSTEADOFQSPAPPL : BOOL;
	XPDOINTERFACEDISABLED : BOOL;
	XPLNOTVALID : BOOL;
	XPPIACTIVE : BOOL;
	XMAGNETISATIONFINISHED : BOOL;
	XFAULTACTIVE : BOOL;
	XFAULTREACTIONACTIVE : BOOL;
	XFIRSTERRORCYCLE : BOOL;
	XWARNINGACTIVE : BOOL;
	WTEXTREFID : WORD;
	DWDRIVEERRORID : DWORD;
	XSERVICEMODEHANDLINGINDRIVEACTIVE : BOOL;
	XBRAKESTATUSBIT : BOOL;
	XSBCACTIVE : BOOL;
END_STRUCT
END_TYPE

(* ---- L_MC1P_DRIVETYPE.dut ---- *)
TYPE L_MC1P_DRIVETYPE :
(
	VIRTUAL := 0,
	HL9400 := 1,
	I700 := 2,
	ENCODER := 3,
	GENERICDRIVE := 4,
	I500 := 5,
	I900 := 6,
	I900DRIVE := 7,
	I750 := 8,
	UNIVERSAL := 10
);
END_TYPE

(* ---- L_MC1P_ENCODERTYPE.dut ---- *)
TYPE L_MC1P_ENCODERTYPE :
(
	UNKNOWN := 0,
	FREEENCODER := 1,
	BPBENCODER := 2,
	I500ECAT := 3,
	I900ENCDRIVE := 4,
	I900ECAT := 5,
	ECATENCODER := 6
);
END_TYPE

(* ---- L_MC1P_ERRORINFORMATION.dut ---- *)
TYPE L_MC1P_ERRORINFORMATION :
STRUCT
	EERRORID : L_IE1P_Error;
	XWARNING : BOOL;
	PINSTANCE : DWORD := 0;
	TTIMESTAMP : TIME;
	TRESETTIMESTAMP : TIME;
	DWEXTENDEDERRORINFO : DWORD;
	PSINSTANCENAME : POINTER TO STRING;
END_STRUCT
END_TYPE

(* ---- L_MC1P_EXECUTIONINDEX.dut ---- *)
TYPE L_MC1P_EXECUTIONINDEX :
(
	FIRST := 1,
	SECOND := 2
);
END_TYPE

(* ---- L_MC1P_FASTOUTPUTINPUT.dut ---- *)
TYPE L_MC1P_FASTOUTPUTINPUT :
STRUCT
	XEXECUTE : BOOL;
	XABORT : BOOL;
	BYDIGITALOUTPUTSEL : BYTE := 1;
	XOUTPUTSTATE : BOOL;
	LRSWITCHPOSITION : LREAL;
	WEXTERNALDELAYCOMPENSATION : WORD;
	LRDYNVELPOSOFFSET : LREAL;
	XRESET : BOOL;
	XDISABLEACCCALC : BOOL := FALSE;
	EVALUESOURCE : MC_SOURCE := MC_SOURCE.mcActualValue;
END_STRUCT
END_TYPE

(* ---- L_MC1P_FASTOUTPUTOUTPUT.dut ---- *)
TYPE L_MC1P_FASTOUTPUTOUTPUT :
STRUCT
	XDONE : BOOL;
	XBUSY : BOOL;
	XCOMMANDABORTED : BOOL;
	XERROR : BOOL;
	EERRORID : L_IE1P_Error;
END_STRUCT
END_TYPE

(* ---- L_MC1P_FOLLOWSETVALUESINPUT.dut ---- *)
TYPE L_MC1P_FOLLOWSETVALUESINPUT :
STRUCT
	XCONTINUOUSUPDATE : BOOL := TRUE;
	LRPOSITION : LREAL;
	LRVELOCITY : LREAL := 0;
	LRACCELERATION : LREAL := 0;
	ESETVALUEMODE : L_MC1P_SetValueMode := L_MC1P_SetValueMode.Pos;
	LRPOSDIFFIN : LREAL;
END_STRUCT
END_TYPE

(* ---- L_MC1P_FOLLOWSETVALUESOUTPUT.dut ---- *)
TYPE L_MC1P_FOLLOWSETVALUESOUTPUT :
STRUCT
END_STRUCT
END_TYPE

(* ---- L_MC1P_FORCESETVALUESINPUT.dut ---- *)
TYPE L_MC1P_FORCESETVALUESINPUT :
STRUCT
	LRFORCEDPOSITION : LREAL;
	LRFORCEDVELOCITY : LREAL;
	LRFORCEDACCELERATION : LREAL;
	LRFORCEDTORQUE : LREAL;
END_STRUCT
END_TYPE

(* ---- L_MC1P_FORCESETVALUESOUTPUT.dut ---- *)
TYPE L_MC1P_FORCESETVALUESOUTPUT :
STRUCT
END_STRUCT
END_TYPE

(* ---- L_MC1P_GETMAXVELACCDECINPUT.dut ---- *)
TYPE L_MC1P_GETMAXVELACCDECINPUT :
STRUCT
	XENABLE : BOOL;
	DWTIMESTAMP : DWORD;
	EMC_SOURCE : MC_SOURCE;
END_STRUCT
END_TYPE

(* ---- L_MC1P_GETMAXVELACCDECOUTPUT.dut ---- *)
TYPE L_MC1P_GETMAXVELACCDECOUTPUT :
STRUCT
	XVALID : BOOL;
	XBUSY : BOOL;
	XERROR : BOOL;
	EERRORID : L_IE1P_Error;
	LRMAXVELOCITIY : LREAL;
	DWTIMEVELATMAX : DWORD;
	LRMAXACCELERATION : LREAL;
	DWTIMEACCATMAX : DWORD;
	LRMAXDECELERATION : LREAL;
	DWTIMEDECATMAX : DWORD;
END_STRUCT
END_TYPE

(* ---- L_MC1P_GISEQUENCE_EXFAN_LIMITS.dut ---- *)
TYPE L_MC1P_GISEQUENCE_EXFAN_LIMITS :
(
	EGI_EXFAN_LIMITS_INIT,
	EGI_EXFAN_LIMITS_FIRSTRAMP,
	EGI_EXFAN_LIMITS_SECONDRAMP,
	EGI_EXFAN_LIMITS_GENERATEPULSE,
	EGI_EXFAN_LIMITS_CHECKDISTANCE,
	EGI_EXFAN_LIMITS_CALCULATEMOVETIME,
	EGI_EXFAN_LIMITS_MOVETOLIMIT
);
END_TYPE

(* ---- L_MC1P_GISEQUENCE_EXFAN_NOLIMITS.dut ---- *)
TYPE L_MC1P_GISEQUENCE_EXFAN_NOLIMITS :
(
	EGI_EXFAN_NOLIMITS_INIT,
	EGI_EXFAN_NOLIMITS_FIRSTRAMP,
	EGI_EXFAN_NOLIMITS_SECONDRAMP,
	EGI_EXFAN_NOLIMITS_GENERATEPULSE,
	EGI_EXFAN_NOLIMITS_CHECKDIRECTION
);
END_TYPE

(* ---- L_MC1P_GISEQUENCE_NOEXFAN_LIMITS.dut ---- *)
TYPE L_MC1P_GISEQUENCE_NOEXFAN_LIMITS :
(
	EGI_NOEXFAN_LIMITS_INIT,
	EGI_NOEXFAN_LIMITS_FIRSTRAMP,
	EGI_NOEXFAN_LIMITS_SECONDRAMP,
	EGI_NOEXFAN_LIMITS_GENERATEPULSE,
	EGI_NOEXFAN_LIMITS_WAITONTIME,
	EGI_NOEXFAN_LIMITS_CHECKDISTANCE,
	EGI_NOEXFAN_LIMITS_CALCULATEMOVETIME,
	EGI_NOEXFAN_LIMITS_MOVETOLIMIT
);
END_TYPE

(* ---- L_MC1P_GISEQUENCE_NOEXFAN_NOLIMITS.dut ---- *)
TYPE L_MC1P_GISEQUENCE_NOEXFAN_NOLIMITS :
(
	EGI_NOEXFAN_NOLIMITS_INIT,
	EGI_NOEXFAN_NOLIMITS_FIRSTRAMP,
	EGI_NOEXFAN_NOLIMITS_GENERATEPULSE,
	EGI_NOEXFAN_NOLIMITS_WAITONTIME,
	EGI_NOEXFAN_NOLIMITS_CHECKDIRECTION
);
END_TYPE

(* ---- L_MC1P_GRINDINMODE.dut ---- *)
TYPE L_MC1P_GRINDINMODE :
(
	CW := 1,
	CCW := 2,
	CWCCW := 3,
	CCWCW := 4
);
END_TYPE

(* ---- L_MC1P_GRINDINSEQUENCE.dut ---- *)
TYPE L_MC1P_GRINDINSEQUENCE :
(
	EGI_DEFAULT := 0,
	EGI_INIT,
	EGI_CONTROLMODE,
	EGI_RAMP1,
	EGI_RAMP2,
	EGI_RAMPDOWN,
	EGI_PULS1,
	EGI_PULS2,
	EGI_DISABLE,
	EGI_CHOOSESTEPSEQUENCE,
	EGI_CALLSTEPSEQUENCE1,
	EGI_CALLSTEPSEQUENCE2,
	EGI_CALLSTEPSEQUENCE3,
	EGI_CALLSTEPSEQUENCE4,
	EGI_CALCULATEDOWNRAMPTYPE,
	EGI_DONE
);
END_TYPE

(* ---- L_MC1P_HALTINPUT.dut ---- *)
TYPE L_MC1P_HALTINPUT :
STRUCT
	EXECUTE : BOOL;
	DECELERATION : LREAL;
	JERK : LREAL;
	BUFFERMODE : MC_BUFFER_MODE;
	CALLEDBYABC : BOOL;
	CONTINUOUSUPDATE : BOOL;
END_STRUCT
END_TYPE

(* ---- L_MC1P_HALTOUTPUT.dut ---- *)
TYPE L_MC1P_HALTOUTPUT :
STRUCT
	DONE : BOOL;
	BUSY : BOOL;
	ACTIVE : BOOL;
	COMMANDABORTED : BOOL;
	ERROR : BOOL;
	ERRORID : L_IE1P_Error;
	XUSED : BOOL;
END_STRUCT
END_TYPE

(* ---- L_MC1P_HALTSUPERIMPOSEDINPUT.dut ---- *)
TYPE L_MC1P_HALTSUPERIMPOSEDINPUT :
STRUCT
	EXECUTE : BOOL;
	DECELERATION : LREAL;
	JERK : LREAL;
END_STRUCT
END_TYPE

(* ---- L_MC1P_HALTSUPERIMPOSEDOUTPUT.dut ---- *)
TYPE L_MC1P_HALTSUPERIMPOSEDOUTPUT :
STRUCT
	DONE : BOOL;
	BUSY : BOOL;
	ACTIVE : BOOL;
	COMMANDABORTED : BOOL;
	ERROR : BOOL;
	ERRORID : L_IE1P_Error;
END_STRUCT
END_TYPE

(* ---- L_MC1P_HOMEINPUT.dut ---- *)
TYPE L_MC1P_HOMEINPUT :
STRUCT
	EXECUTE : BOOL;
	POSITION : LREAL;
	BUFFERMODE : MC_BUFFER_MODE;
	HOMEABSSWITCH : BOOL;
	USEEXTPARAMETER : BOOL;
	EXTPARAMETER : L_MC1P_HomeParameter;
	EXTTP : MC_TRIGGER_REF;
	USEPOSITIONINPUT : BOOL := TRUE;
END_STRUCT
END_TYPE

(* ---- L_MC1P_HOMEMODE.dut ---- *)
TYPE L_MC1P_HOMEMODE :
(
	CWTORQUELIMIT := -2,
	CCWTORQUELIMIT := -1,
	SETPOSITIONDIRECT := 0,
	CCWLIMITSWITCHCWTP := 1,
	CWLIMITSWITCHCCWTP := 2,
	CWRPCCWRNTP := 3,
	CCWRPCWRNTP := 5,
	CCWLIMITSWITCH := 17,
	CWLIMITSWITCH := 18,
	CWRPCCWRN := 19,
	CCWRPCWRN := 21,
	CCWTP := 33,
	CWTP := 34,
	SETPOSITIONINANYSTATE := 97,
	SETOFFSETINANYSTATE := 98,
	RESETHOMEINFO := 99,
	DRIVEBASED := 100
);
END_TYPE

(* ---- L_MC1P_HOMEOUTPUT.dut ---- *)
TYPE L_MC1P_HOMEOUTPUT :
STRUCT
	DONE : BOOL;
	BUSY : BOOL;
	ACTIVE : BOOL;
	COMMANDABORTED : BOOL;
	ERROR : BOOL;
	ERRORID : L_IE1P_Error;
	XUSED : BOOL;
END_STRUCT
END_TYPE

(* ---- L_MC1P_HOMEPARAMETER.dut ---- *)
TYPE L_MC1P_HOMEPARAMETER :
STRUCT
	EHOMEMODE : L_MC1P_HomeMode;
	EHOMESTOPMODE : L_MC1P_HomeStopMode;
	LRTARGETPOSITION : LREAL;
	LRVELOCITY1 : LREAL;
	LRVELOCITY2 : LREAL;
	LRACCELERATION1 : LREAL;
	LRACCELERATION2 : LREAL;
	LRJERK : LREAL;
	RTORQUELIMIT : REAL;
	RTORQUETIME : REAL;
	DWTPCONFIG : L_MC1P_HomeTPMode;
	WDRIVEHOMEMODE : WORD;
	ESTOPMODEDIRECTION : MC_DIRECTION;
	LROFFSETPOSITION : LREAL;
END_STRUCT
END_TYPE

(* ---- L_MC1P_HOMESTOPMODE.dut ---- *)
TYPE L_MC1P_HOMESTOPMODE :
(
	STOPPOSITIONING := 0,
	RELATIVEPOSITIONING := 1,
	ABSOLUTEPOSITIONING := 2
);
END_TYPE

(* ---- L_MC1P_HOMETPMODE.dut ---- *)
TYPE L_MC1P_HOMETPMODE :
(
	EXTERNALSOURCE := 0,
	TP1_POSEDGE := 1,
	TP1_NEGEDGE := 2,
	TP1_ANYEDGE := 3,
	TP1_ZEROPULSE := 4,
	TP1_ZEROPULSE2NDFDB := 5,
	TP2_POSEDGE := 11,
	TP2_NEGEDGE := 12,
	TP2_ANYEDGE := 13,
	TP2_ZEROPULSE := 14,
	TP2_ZEROPULSEFDB2ND := 15,
	TP3_POSEDGE := 21,
	TP3_NEGEDGE := 22,
	TP3_ANYEDGE := 23,
	TP3_ZEROPULSE := 24,
	TP3_ZEROPULSEFDB2ND := 25,
	TP4_POSEDGE := 31,
	TP4_NEGEDGE := 32,
	TP4_ANYEDGE := 33,
	TP4_ZEROPULSE := 34,
	TP5_ZEROPULSEFDB2ND := 35
);
END_TYPE

(* ---- L_MC1P_HWLIMITSWITCHINTERFACEINPUT.dut ---- *)
TYPE L_MC1P_HWLIMITSWITCHINTERFACEINPUT :
STRUCT
	XENABLE : BOOL;
	XLIMITSWITCHPOS : BOOL;
	XLIMITSWITCHNEG : BOOL;
	XOVERWRITEOTHERSOURCES : BOOL;
	XHOMEABSSWITCH : BOOL;
END_STRUCT
END_TYPE

(* ---- L_MC1P_HWLIMITSWITCHINTERFACEOUTPUT.dut ---- *)
TYPE L_MC1P_HWLIMITSWITCHINTERFACEOUTPUT :
STRUCT
	XBUSY : BOOL;
	XERROR : BOOL;
	EERRORID : L_IE1P_Error;
END_STRUCT
END_TYPE

(* ---- L_MC1P_I900REFOFFSETHANDLING.dut ---- *)
TYPE L_MC1P_I900REFOFFSETHANDLING :
STRUCT
	DWSWITCHCYCLECOUNTER : DWORD;
	DIDRIVEREFOFFSET : DINT;
END_STRUCT
END_TYPE

(* ---- L_MC1P_INTERFACEID.dut ---- *)
TYPE L_MC1P_INTERFACEID :
(
	L_MC1P_ITOUCHPROBEHANDLER := (L_MC1P_Internal.cdiEnumStartValue + 1),
	L_MC1P_IAXIS_REF_MASTERVALUES := (L_MC1P_Internal.cdiEnumStartValue + 2)
);
END_TYPE

(* ---- L_MC1P_INTERNALBRAKEMODE.dut ---- *)
TYPE L_MC1P_INTERNALBRAKEMODE :
(
	BM_OFF := 0,
	BM_MANINT := 11,
	BM_AUTINT := 12,
	BM_MANEXT := 1,
	BM_AUTEXT := 2,
	BM_AUTGSB := 22
);
END_TYPE

(* ---- L_MC1P_INTERPOLATIONMODE.dut ---- *)
TYPE L_MC1P_INTERPOLATIONMODE :
(
	LINEAR := 0,
	QUADRATICPOS := 1
);
END_TYPE

(* ---- L_MC1P_INTPROFILEDATA.dut ---- *)
TYPE L_MC1P_INTPROFILEDATA :
STRUCT
	PHASE1 : L_MC1P_ProfilePhaseData;
	PHASE2 : L_MC1P_ProfilePhaseData;
	PHASE3 : L_MC1P_ProfilePhaseData;
	PHASE4 : L_MC1P_ProfilePhaseData;
	PHASE5 : L_MC1P_ProfilePhaseData;
	PHASE6 : L_MC1P_ProfilePhaseData;
	PHASE7 : L_MC1P_ProfilePhaseData;
END_STRUCT
END_TYPE

(* ---- L_MC1P_INTPROFILEDATAACC.dut ---- *)
TYPE L_MC1P_INTPROFILEDATAACC :
STRUCT
	PHASE1 : L_MC1P_ProfilePhaseData;
	PHASE2 : L_MC1P_ProfilePhaseData;
	PHASE3 : L_MC1P_ProfilePhaseData;
END_STRUCT
END_TYPE

(* ---- L_MC1P_KINDOFMOTION.dut ---- *)
TYPE L_MC1P_KINDOFMOTION :
(
	NOTDEFINED := 0,
	TRANSLATORY := 1,
	ROTARY := 2
);
END_TYPE

(* ---- L_MC1P_LIMITERINPUT_INTERNAL.dut ---- *)
TYPE L_MC1P_LIMITERINPUT_INTERNAL :
STRUCT
	PAXIS : POINTER TO AXIS_REF;
	XENABLE : BOOL;
	DWLIMITERCONTROL : DWORD;
END_STRUCT
END_TYPE

(* ---- L_MC1P_LIMITEROUTPUT_INTERNAL.dut ---- *)
TYPE L_MC1P_LIMITEROUTPUT_INTERNAL :
STRUCT
	XBUSY : BOOL;
	XERROR : BOOL;
	EERRORID : L_IE1P_Error;
	DWSTATE : DWORD;
	XLIMITATIONACTIVE : BOOL;
	XSLSACTIVE : BOOL;
	LRACTLIMITEDVELOCITY : LREAL;
	LRACTLIMITEDDECTIME : LREAL;
	LRACTLIMITEDJERK : LREAL;
END_STRUCT
END_TYPE

(* ---- L_MC1P_MANIPULATIONBASEINPUT.dut ---- *)
TYPE L_MC1P_MANIPULATIONBASEINPUT :
STRUCT
	XENABLE : BOOL;
	EEXECUTIONINDEX : L_MC1P_ExecutionIndex := L_MC1P_ExecutionIndex.First;
	XIGNOREFILTERONSTOP : BOOL;
END_STRUCT
END_TYPE

(* ---- L_MC1P_MANIPULATIONBASEOUTPUT.dut ---- *)
TYPE L_MC1P_MANIPULATIONBASEOUTPUT :
STRUCT
	XBUSY : BOOL;
	XACTIVE : BOOL;
	XERROR : BOOL;
	EERRORID : L_IE1P.L_IE1P_Error;
	LRSETPOSOUT : LREAL;
	LRSETVELOUT : LREAL;
	LRSETACCOUT : LREAL;
	LRSETTORQUEOUT : LREAL;
END_STRUCT
END_TYPE

(* ---- L_MC1P_MANJOGOPENLOOPINPUT.dut ---- *)
TYPE L_MC1P_MANJOGOPENLOOPINPUT :
STRUCT
	XENABLE : BOOL;
	XJOGPOSITIVE : BOOL;
	XJOGNEGATIVE : BOOL;
	XPARAMETERSET2 : BOOL;
END_STRUCT
END_TYPE

(* ---- L_MC1P_MANJOGOPENLOOPOUTPUT.dut ---- *)
TYPE L_MC1P_MANJOGOPENLOOPOUTPUT :
STRUCT
	XBUSY : BOOL;
	XOPERATIONENABLED : BOOL;
	XDONE : BOOL;
	XACTIVE : BOOL;
	XCOMMANDABORTED : BOOL;
	XERROR : BOOL;
	EERRORID : L_IE1P_Error;
END_STRUCT
END_TYPE

(* ---- L_MC1P_MANUALJOGINPUT_INTERNAL.dut ---- *)
TYPE L_MC1P_MANUALJOGINPUT_INTERNAL :
STRUCT
	PAXIS : POINTER TO AXIS_REF;
	XJOGPOSITIVE : BOOL;
	XJOGNEGATIVE : BOOL;
	XCONTINUOUSUPDATE : BOOL;
	LRVELOCITY : LREAL;
	LRACCELERATION : LREAL;
	LRDECELERATION : LREAL;
	LRJERK : LREAL;
	LRJERKDEC : LREAL;
	XSTEPMODE : BOOL;
	LRDISTANCE : LREAL;
END_STRUCT
END_TYPE

(* ---- L_MC1P_MANUALJOGOUTPUT_INTERNAL.dut ---- *)
TYPE L_MC1P_MANUALJOGOUTPUT_INTERNAL :
STRUCT
	XBUSY : BOOL;
	XDONE : BOOL;
	XCOMMANDABORTED : BOOL;
	XERROR : BOOL;
	EERRORID : L_IE1P_Error;
	XUSED : BOOL;
END_STRUCT
END_TYPE

(* ---- L_MC1P_MAPPEDELEMENT.dut ---- *)
TYPE L_MC1P_MAPPEDELEMENT :
STRUCT
	WPARAMETER : WORD;
	WSIZE : WORD;
	PBADRESS : POINTER TO BYTE;
	PADDITIONALDATA : POINTER TO BYTE;
END_STRUCT
END_TYPE

(* ---- L_MC1P_MAPPEDOBJECTS.dut ---- *)
TYPE L_MC1P_MAPPEDOBJECTS :
STRUCT
	INDEXSUBINDEX : DWORD;
	USISIZE : USINT;
	XUSEDBYAXISREF : BOOL;
	PDATA : POINTER TO BYTE;
END_STRUCT
END_TYPE

(* ---- L_MC1P_MCTRLCONTROL.dut ---- *)
TYPE L_MC1P_MCTRLCONTROL :
(
	MCSTANDARD := 0,
	MCUF := 4,
	MCFTC := 5
);
END_TYPE

(* ---- L_MC1P_MEASUREDISTANCEINPUT.dut ---- *)
TYPE L_MC1P_MEASUREDISTANCEINPUT :
STRUCT
	XENABLE : BOOL;
	EMC_SOURCE : MC_SOURCE;
END_STRUCT
END_TYPE

(* ---- L_MC1P_MEASUREDISTANCEOUTPUT.dut ---- *)
TYPE L_MC1P_MEASUREDISTANCEOUTPUT :
STRUCT
	XVALID : BOOL;
	XBUSY : BOOL;
	XERROR : BOOL;
	EERRORID : L_IE1P_Error;
	LRDISTANCE : LREAL;
END_STRUCT
END_TYPE

(* ---- L_MC1P_MINMAXVALUE.dut ---- *)
TYPE L_MC1P_MINMAXVALUE :
STRUCT
	LRMIN : LREAL := 0;
	LRMAX : LREAL := 0;
END_STRUCT
END_TYPE

(* ---- L_MC1P_MOLSTATE.dut ---- *)
TYPE L_MC1P_MOLSTATE :
(
	IDLE := 0,
	CHECKMOLACTIVATION := 1,
	MOLCYCLIC := 2,
	ERROR := 999
);
END_TYPE

(* ---- L_MC1P_MOVEABSOLUTEINPUT_INTERNAL.dut ---- *)
TYPE L_MC1P_MOVEABSOLUTEINPUT_INTERNAL :
STRUCT
	PAXIS : POINTER TO AXIS_REF;
	EXECUTE : BOOL;
	CONTINUOUSUPDATE : BOOL;
	POSITION : LREAL;
	VELOCITY : LREAL;
	ACCELERATION : LREAL;
	DECELERATION : LREAL;
	JERK : LREAL;
	JERKDEC : LREAL;
	DIRECTION : MC_DIRECTION;
	BUFFERMODE : MC_BUFFER_MODE;
END_STRUCT
END_TYPE

(* ---- L_MC1P_MOVEABSOLUTEOUTPUT_INTERNAL.dut ---- *)
TYPE L_MC1P_MOVEABSOLUTEOUTPUT_INTERNAL :
STRUCT
	DONE : BOOL;
	BUSY : BOOL;
	ACTIVE : BOOL;
	COMMANDABORTED : BOOL;
	ERROR : BOOL;
	ERRORID : L_IE1P_Error;
	XUSED : BOOL;
END_STRUCT
END_TYPE

(* ---- L_MC1P_MOVEADDITIVEINPUT.dut ---- *)
TYPE L_MC1P_MOVEADDITIVEINPUT :
STRUCT
	EXECUTE : BOOL;
	CONTINUOUSUPDATE : BOOL;
	DISTANCE : LREAL;
	VELOCITY : LREAL;
	ACCELERATION : LREAL;
	DECELERATION : LREAL;
	JERK : LREAL;
	BUFFERMODE : MC_BUFFER_MODE;
	JERKDEC : LREAL;
END_STRUCT
END_TYPE

(* ---- L_MC1P_MOVEADDITIVEOUTPUT.dut ---- *)
TYPE L_MC1P_MOVEADDITIVEOUTPUT :
STRUCT
	DONE : BOOL;
	BUSY : BOOL;
	ACTIVE : BOOL;
	COMMANDABORTED : BOOL;
	ERROR : BOOL;
	ERRORID : L_IE1P_Error;
END_STRUCT
END_TYPE

(* ---- L_MC1P_MOVECONTINUOUSABSOLUTEINPUT.dut ---- *)
TYPE L_MC1P_MOVECONTINUOUSABSOLUTEINPUT :
STRUCT
	EXECUTE : BOOL;
	CONTINUOUSUPDATE : BOOL;
	POSITION : LREAL;
	ENDVELOCITY : LREAL;
	VELOCITY : LREAL;
	ACCELERATION : LREAL;
	DECELERATION : LREAL;
	JERK : LREAL;
	DIRECTION : MC_DIRECTION;
	BUFFERMODE : MC_BUFFER_MODE;
	JERKDEC : LREAL;
END_STRUCT
END_TYPE

(* ---- L_MC1P_MOVECONTINUOUSABSOLUTEOUTPUT.dut ---- *)
TYPE L_MC1P_MOVECONTINUOUSABSOLUTEOUTPUT :
STRUCT
	INENDVELOCITY : BOOL;
	BUSY : BOOL;
	ACTIVE : BOOL;
	COMMANDABORTED : BOOL;
	ERROR : BOOL;
	ERRORID : L_IE1P_Error;
END_STRUCT
END_TYPE

(* ---- L_MC1P_MOVECONTINUOUSRELATIVEINPUT.dut ---- *)
TYPE L_MC1P_MOVECONTINUOUSRELATIVEINPUT :
STRUCT
	EXECUTE : BOOL;
	CONTINUOUSUPDATE : BOOL;
	DISTANCE : LREAL;
	ENDVELOCITY : LREAL;
	VELOCITY : LREAL;
	ACCELERATION : LREAL;
	DECELERATION : LREAL;
	JERK : LREAL;
	BUFFERMODE : MC_BUFFER_MODE;
	JERKDEC : LREAL;
END_STRUCT
END_TYPE

(* ---- L_MC1P_MOVECONTINUOUSRELATIVEOUTPUT.dut ---- *)
TYPE L_MC1P_MOVECONTINUOUSRELATIVEOUTPUT :
STRUCT
	INENDVELOCITY : BOOL;
	BUSY : BOOL;
	ACTIVE : BOOL;
	COMMANDABORTED : BOOL;
	ERROR : BOOL;
	ERRORID : L_IE1P_Error;
END_STRUCT
END_TYPE

(* ---- L_MC1P_MOVERELATIVEINPUT.dut ---- *)
TYPE L_MC1P_MOVERELATIVEINPUT :
STRUCT
	EXECUTE : BOOL;
	CONTINUOUSUPDATE : BOOL;
	DISTANCE : LREAL;
	VELOCITY : LREAL;
	ACCELERATION : LREAL;
	DECELERATION : LREAL;
	JERK : LREAL;
	JERKDEC : LREAL;
	BUFFERMODE : MC_BUFFER_MODE;
	XUSEEXTERNPROFILECALCULATION : BOOL;
	ITFPOSPROFILECALCULATION : L_MC1P_IPosProfileCalculation;
END_STRUCT
END_TYPE

(* ---- L_MC1P_MOVERELATIVEOUTPUT.dut ---- *)
TYPE L_MC1P_MOVERELATIVEOUTPUT :
STRUCT
	DONE : BOOL;
	BUSY : BOOL;
	ACTIVE : BOOL;
	COMMANDABORTED : BOOL;
	ERROR : BOOL;
	ERRORID : L_IE1P_Error;
	XUSED : BOOL;
END_STRUCT
END_TYPE

(* ---- L_MC1P_MOVESUPERIMPOSEDINPUT.dut ---- *)
TYPE L_MC1P_MOVESUPERIMPOSEDINPUT :
STRUCT
	EXECUTE : BOOL;
	CONTINUOUSUPDATE : BOOL;
	DISTANCE : LREAL;
	VELOCITYDIFF : LREAL;
	ACCELERATION : LREAL;
	DECELERATION : LREAL;
	JERK : LREAL;
	JERKDEC : LREAL;
END_STRUCT
END_TYPE

(* ---- L_MC1P_MOVESUPERIMPOSEDOUTPUT.dut ---- *)
TYPE L_MC1P_MOVESUPERIMPOSEDOUTPUT :
STRUCT
	DONE : BOOL;
	BUSY : BOOL;
	ACTIVE : BOOL;
	COMMANDABORTED : BOOL;
	ERROR : BOOL;
	ERRORID : L_IE1P_Error;
	COVEREDDISTANCE : LREAL;
END_STRUCT
END_TYPE

(* ---- L_MC1P_MOVEVELOCITYINPUT.dut ---- *)
TYPE L_MC1P_MOVEVELOCITYINPUT :
STRUCT
	EXECUTE : BOOL;
	CONTINUOUSUPDATE : BOOL;
	POSITION : LREAL;
	VELOCITY : LREAL;
	ACCELERATION : LREAL;
	DECELERATION : LREAL;
	JERK : LREAL;
	JERKDEC : LREAL;
	DIRECTION : MC_DIRECTION;
	BUFFERMODE : MC_BUFFER_MODE;
	XUSEEXTERNPROFILECALCULATION : BOOL;
	ITFPOSPROFILECALCULATION : L_MC1P_IPosProfileCalculation;
	XENABLEOFFSETVELOCITY : BOOL;
	LROFFSETVELOCITY : LREAL;
END_STRUCT
END_TYPE

(* ---- L_MC1P_MOVEVELOCITYOUTPUT.dut ---- *)
TYPE L_MC1P_MOVEVELOCITYOUTPUT :
STRUCT
	INVELOCITY : BOOL;
	BUSY : BOOL;
	ACTIVE : BOOL;
	COMMANDABORTED : BOOL;
	ERROR : BOOL;
	ERRORID : L_IE1P_Error;
	XUSED : BOOL;
END_STRUCT
END_TYPE

(* ---- L_MC1P_MULTIAXISINFO.dut ---- *)
TYPE L_MC1P_MULTIAXISINFO :
STRUCT
	UIDEVICESLOT : UINT;
	UIOFFSETDRIVEPARA : UINT;
	ITFSLAVEMULTIAXISMODULEHANDLER : L_IMHP_IModuleHandler;
	ITFSLAVEAXISMODULEHANDLER : L_IMHP_IModuleHandler;
END_STRUCT
END_TYPE

(* ---- L_MC1P_OPTICALTRACKINGINPUT.dut ---- *)
TYPE L_MC1P_OPTICALTRACKINGINPUT :
STRUCT
	XEXECUTE : BOOL := FALSE;
	RTIME : REAL := 5.0;
END_STRUCT
END_TYPE

(* ---- L_MC1P_OPTICALTRACKINGOUTPUT.dut ---- *)
TYPE L_MC1P_OPTICALTRACKINGOUTPUT :
STRUCT
	XDONE : BOOL := FALSE;
	XBUSY : BOOL;
	XERROR : BOOL;
	EERRORID : L_IE1P_Error;
END_STRUCT
END_TYPE

(* ---- L_MC1P_ORDINALTYPE.dut ---- *)
TYPE L_MC1P_ORDINALTYPE :
(
	OTNONE := 0,
	OTBOOL := 1,
	OTBYTE := 2,
	OTSINT := 3,
	OTUSINT := 4,
	OTWORD := 5,
	OTINT := 6,
	OTUINT := 7,
	OTDWORD := 8,
	OTDINT := 9,
	OTUDINT := 10,
	OTLWORD := 11,
	OTLINT := 12,
	OTULINT := 13,
	OTREAL := 14,
	OTLREAL := 15
);
END_TYPE

(* ---- L_MC1P_PARACCESS.dut ---- *)
TYPE L_MC1P_PARACCESS :
STRUCT
	AXISNAME : REFERENCE TO STRING;
	DEVICETYPE : REFERENCE TO WORD;
	AXISSTATE : REFERENCE TO WORD;
	AXISSTATUSWORD : REFERENCE TO DWORD;
	ACTIVEERRORID : REFERENCE TO WORD;
	AXISCONTROLWORD : REFERENCE TO WORD;
	AXISCONFIGURATION : REFERENCE TO DWORD;
	ACTPOSITION : REFERENCE TO LREAL;
	ACTVELOCITY : REFERENCE TO LREAL;
	ACTACCELERATION : REFERENCE TO LREAL;
	ACTTORQUE : REFERENCE TO LREAL;
	SETPOSITION : REFERENCE TO LREAL;
	SETVELOCITY : REFERENCE TO LREAL;
	SETACCELERATION : REFERENCE TO LREAL;
	SETTORQUE : REFERENCE TO LREAL;
	KINDOFMOTIONSELECTION : REFERENCE TO WORD;
	ACTIVEUNIT : REFERENCE TO WORD;
	RATIONUMERATORADD : REFERENCE TO DWORD;
	RATIODENOMINATORADD : REFERENCE TO DWORD;
	AXISMODE : REFERENCE TO WORD;
	UDITOTALMEASURINGRANGE : REFERENCE TO UDINT;
	USEASVIRTUAL : REFERENCE TO BOOL;
	TRAVERSINGRANGE : REFERENCE TO WORD;
	CYCLELENGTH : REFERENCE TO LREAL;
	FEEDCONSTANT : REFERENCE TO LREAL;
	RATIONUMERATOR : REFERENCE TO DWORD;
	RATIODENOMINATOR : REFERENCE TO DWORD;
	ORIENTATIONINV : REFERENCE TO BOOL;
	INKPERREV : REFERENCE TO DWORD;
	INERTIALOAD : REFERENCE TO LREAL;
	INERTIAMOTOR : REFERENCE TO LREAL;
	REFTORQUE : REFERENCE TO LREAL;
	DEFAULTVELOCITY : REFERENCE TO LREAL;
	DEFAULTACCELERATION : REFERENCE TO LREAL;
	DEFAULTJERK : REFERENCE TO LREAL;
	MOTORRATEDVELOCITY : REFERENCE TO LREAL;
	MAXVELOCITY : REFERENCE TO LREAL;
	MAXACCELERATION : REFERENCE TO LREAL;
	MAXJERK : REFERENCE TO LREAL;
	DECERRORSTOP : REFERENCE TO LREAL;
	JERKERRORSTOP : REFERENCE TO LREAL;
	ENABLESWLIMIT : REFERENCE TO BOOL;
	SWLIMITPOS : REFERENCE TO LREAL;
	SWLIMITNEG : REFERENCE TO LREAL;
	BEHAVEONSWLIMIT : REFERENCE TO WORD;
	ENABLEFOLLOWINGERROR : REFERENCE TO BOOL;
	MAXFOLLOWINGERRORWARNING : REFERENCE TO LREAL;
	MAXFOLLOWINGERRORERROR : REFERENCE TO LREAL;
	ACTFOLLOWINGERROR : REFERENCE TO LREAL;
	MAXFOLLOWINGERROR : REFERENCE TO LREAL;
	FOLLOWINGERRORREACTION : REFERENCE TO WORD;
	ENCODERINPUTFILTER : REFERENCE TO USINT;
	ENCODERPOSFILTERSTATE : REFERENCE TO WORD;
	ENCODERVELFILTERSTATE : REFERENCE TO WORD;
	BTWFILTERTIME : REFERENCE TO DINT;
	REDPOSQUANT : REFERENCE TO WORD;
	ENCFILTERCYCLES : REFERENCE TO WORD;
	ENCFILTERCYCLESPOS : REFERENCE TO WORD;
	COMPENSATIONMODE : REFERENCE TO WORD;
	SETVALDELAYTIME : REFERENCE TO LREAL;
	ENCODERUPDATETIME : REFERENCE TO DWORD;
	HOMING_MODE : REFERENCE TO INT;
	HOMING_STOPMODE : REFERENCE TO INT;
	HOMING_TARGETPOSITION : REFERENCE TO LREAL;
	HOMING_VELOCITY1 : REFERENCE TO LREAL;
	HOMING_VELOCITY2 : REFERENCE TO LREAL;
	HOMING_ACCELERATION1 : REFERENCE TO LREAL;
	HOMING_ACCELERATION2 : REFERENCE TO LREAL;
	HOMING_JERK : REFERENCE TO LREAL;
	HOMING_TORQUELIMIT : REFERENCE TO REAL;
	HOMING_TORQUETIME : REFERENCE TO REAL;
	HOMING_TPCONFIG : REFERENCE TO DWORD;
	HOMING_RESTOREHOMEPOSITION : REFERENCE TO BOOL;
	HOMING_RESTORETRESHOLD : REFERENCE TO LREAL;
	HOMING_DRIVEHOMEMODE : REFERENCE TO WORD;
	HOMING_HOMEPOSITION : REFERENCE TO LREAL;
	HOMING_POSSETPERMANENTLY : REFERENCE TO USINT;
	HOMIN_OFFSETPOSITION : REFERENCE TO LREAL;
	HOMING_STOPMODEDIRECTION : REFERENCE TO INT;
	HOMESENSORDISTANCE : REFERENCE TO LREAL;
	CONTROLMODEDEFAULT : REFERENCE TO WORD;
	ACTCONTROLMODE : REFERENCE TO WORD;
	ENCODERNAME : REFERENCE TO STRING;
	POSCTRLGAIN : REFERENCE TO LREAL;
	POSCTRLOUTPUTLIMITATION : REFERENCE TO LREAL;
	POSCTRKOUTPUT : REFERENCE TO LREAL;
	POSCTRLADAPTVALUE : REFERENCE TO UINT;
	POSCTRLADAPTIONFROM0X2985 : REFERENCE TO USINT;
	POSCTRLADAPTACTIVEVALUE : REFERENCE TO UINT;
	SETVALUEMONITORING : REFERENCE TO BOOL;
	TIMELIMITSWITCHON : REFERENCE TO REAL;
	REAKTONMCFBERROR : REFERENCE TO BOOL;
	ENABLELOGENTRY : REFERENCE TO BOOL;
	HWLIMITERRORREACTION : REFERENCE TO USINT;
	SWLIMITERRORREACTION : REFERENCE TO USINT;
	LIMITPROFILEERRORREACTION : REFERENCE TO USINT;
	CINHERRORREACTION : REFERENCE TO USINT;
	LIMITERSTOPREACTION : REFERENCE TO USINT;
	REACTIONSSISTATUS1 : REFERENCE TO USINT;
	BRAKE_MODE : REFERENCE TO DWORD;
	BRAKE_RELEASETIME : REFERENCE TO LREAL;
	BRAKE_ACTIVATIONTIME : REFERENCE TO LREAL;
	BRAKE_ACTMODE : REFERENCE TO DWORD;
	BRAKE_SAMPLEDTORQUE : REFERENCE TO LREAL;
	BRAKE_EFFECTIVETORQUE : REFERENCE TO LREAL;
	BRAKETEST_STATE : REFERENCE TO WORD;
	BRAKE_SOURCESTARTVALUE : REFERENCE TO WORD;
	BRAKE_MSTARTVALUE : REFERENCE TO LREAL;
	BRAKE_BRAKERAMPTIME : REFERENCE TO LREAL;
	BRAKE_BRAKEACCDEPENDING : REFERENCE TO BOOL;
	BRAKETEST_CMD : REFERENCE TO USINT;
	BRAKETEST_MODE : REFERENCE TO USINT;
	BRAKETEST_TORQUE : REFERENCE TO DINT;
	BRAKETEST_THRESHOLD : REFERENCE TO INT;
	BRAKETEST_RAMPTIME : REFERENCE TO INT;
	BRAKETEST_HOLDTIME : REFERENCE TO INT;
	BRAKETEST_ACTTRESHOLD : REFERENCE TO INT;
	TORQUELIMHIGH : REFERENCE TO INT;
	TORQUELIMLOW : REFERENCE TO INT;
	WINDOWTARGETREACHED : REFERENCE TO LREAL;
	WINDOWTARGETREACHEDTIME : REFERENCE TO LREAL;
	WINDOWSTANDSTILL : REFERENCE TO LREAL;
	OPTIMIZEDPROFILECALCULATIONMODE : REFERENCE TO UINT;
	MODPOSTOLERANCE : REFERENCE TO LREAL;
	RECOVERYWINDOWPOS : REFERENCE TO LREAL;
	RECOVERYWINDOWNEG : REFERENCE TO LREAL;
	SERVICEDIRECTION : REFERENCE TO WORD;
	BRAKEGRINDIN_CMD : REFERENCE TO USINT;
	BRAKEGRINDIN_MODE : REFERENCE TO USINT;
	BRAKEGRINDIN_CTRL : REFERENCE TO BYTE;
	BRAKEGRINDIN_SPEED : REFERENCE TO INT;
	BRAKEGRINDIN_RAMPTIME : REFERENCE TO INT;
	BRAKEGRINDIN_ONTIME : REFERENCE TO INT;
	BRAKEGRINDIN_OFFTIME : REFERENCE TO INT;
	BRAKEGRINDIN_CYCLES : REFERENCE TO WORD;
	BRAKEGRINDIN_CYCLESOUT : REFERENCE TO WORD;
	BRAKEGRINDIN_STATE : REFERENCE TO WORD;
	LIMITEDVELOCITY1 : REFERENCE TO LREAL;
	LIMITEDDECELERATION1 : REFERENCE TO LREAL;
	LIMITEDVELOCITY2 : REFERENCE TO LREAL;
	LIMITEDDECELERATION2 : REFERENCE TO LREAL;
	LIMITEDVELOCITY3 : REFERENCE TO LREAL;
	LIMITEDDECELERATION3 : REFERENCE TO LREAL;
	LIMITEDVELOCITY4 : REFERENCE TO LREAL;
	LIMITEDDECELERATION4 : REFERENCE TO LREAL;
	LIMITEDDISTANCE : REFERENCE TO LREAL;
	SLSOFFSETVELOCITY : REFERENCE TO LREAL;
	FOLLOWERSLS : REFERENCE TO BOOL;
	LIMITSPEEDCTRLSLS : REFERENCE TO BOOL;
	DISABLESAFETYINTERFACE : REFERENCE TO DWORD;
	REQUESTSAFETYINTERFACE : REFERENCE TO DWORD;
	SLIDISTANCE : REFERENCE TO LREAL;
	BRAKEGRINDIN_POSLIMIT1 : REFERENCE TO LREAL;
	BRAKEGRINDIN_POSLIMIT2 : REFERENCE TO LREAL;
	AUTOTUNING_CMD : REFERENCE TO USINT;
	AT_VELOCITY : REFERENCE TO LREAL;
	AT_ACCELERATION : REFERENCE TO LREAL;
	AT_DISTANCE : REFERENCE TO LREAL;
	AT_CALCULATEDDISTANCE : REFERENCE TO LREAL;
	AT_VPNFACTOR : REFERENCE TO WORD;
	AT_TNNFACTOR : REFERENCE TO WORD;
	AT_STATE : REFERENCE TO WORD;
	AT_VPPFACTOR : REFERENCE TO WORD;
	AT_VPPFACTOREXT : REFERENCE TO WORD;
	AT_WAITINGTIME : REFERENCE TO LREAL;
	JOGGINGSETVEL : REFERENCE TO LREAL;
	JOGGINGSETACC : REFERENCE TO LREAL;
	JOGGINGSETDEC : REFERENCE TO LREAL;
	JOGGINGSETJERK : REFERENCE TO LREAL;
	HALTDEC : REFERENCE TO LREAL;
	HALTJERK : REFERENCE TO LREAL;
END_STRUCT
END_TYPE

(* ---- L_MC1P_PARAMETERDATASIM.dut ---- *)
TYPE L_MC1P_PARAMETERDATASIM :
STRUCT
	WINDEX : WORD;
	BYSUBINDEX : BYTE;
	PVALUE : POINTER TO BYTE;
	BYNROFBYTE : BYTE;
	XSUPPORTED : BOOL;
	XWRITEACCESS : BOOL;
	XAXISOFFSETSUPPORTED : BOOL;
	EFIXTOLREAL : L_MC1P_ScaleFixToLREAL := L_MC1P_ScaleFixToLREAL.None;
END_STRUCT
END_TYPE

(* ---- L_MC1P_PARAMS.dut ---- *)
TYPE L_MC1P_PARAMS :
(
	AXISNAME := 2,
	DEVICETYPE := 3,
	AXISSTATE := 4,
	AXISSTATUSWORD := 5,
	ACTIVEERRORID := 6,
	AXISCONTROLWORD := 8,
	AXISCONFIGURATION := 9,
	ACTPOSITION := 10,
	ACTVELOCITY := 11,
	ACTACCELERATION := 12,
	ACTTORQUE := 13,
	SETPOSITION := 14,
	SETVELOCITY := 15,
	SETACCELERATION := 16,
	SETTORQUE := 17,
	KINDOFMOTIONSELECTION := 20,
	ACTIVEUNIT := 21,
	RATIONUMERATORADD := 25,
	RATIODENOMINATORADD := 26,
	AXISMODE := 27,
	UDITOTALMEASURINGRANGE := 28,
	USEASVIRTUAL := 29,
	TRAVERSINGRANGE := 30,
	CYCLELENGTH := 31,
	FEEDCONSTANT := 32,
	RATIONUMERATOR := 33,
	RATIODENOMINATOR := 34,
	ORIENTATIONINV := 35,
	INKPERREV := 36,
	INERTIALOAD := 37,
	INERTIAMOTOR := 38,
	REFTORQUE := 39,
	DEFAULTVELOCITY := 40,
	DEFAULTACCELERATION := 41,
	DEFAULTJERK := 43,
	MOTORRATEDVELOCITY := 44,
	MAXVELOCITY := 45,
	MAXACCELERATION := 46,
	MAXJERK := 47,
	DECERRORSTOP := 48,
	JERKERRORSTOP := 49,
	ENABLESWLIMIT := 50,
	SWLIMITPOS := 51,
	SWLIMITNEG := 52,
	BEHAVEONSWLIMIT := 53,
	ENABLEFOLLOWINGERROR := 54,
	MAXFOLLOWINGERRORWARNING := 55,
	MAXFOLLOWINGERRORERROR := 56,
	ACTFOLLOWINGERROR := 57,
	MAXFOLLOWINGERROR := 58,
	FOLLOWINGERRORREACTION := 59,
	ENCODERINPUTFILTER := 60,
	ENCODERPOSFILTERSTATE := 61,
	ENCODERVELFILTERSTATE := 62,
	BTWFILTERTIME := 63,
	REDPOSQUANT := 64,
	ENCFILTERCYCLES := 65,
	ENCFILTERCYCLESPOS := 66,
	COMPENSATIONMODE := 67,
	SETVALDELAYTIME := 68,
	ENCODERUPDATETIME := 69,
	HOMING_MODE := 70,
	HOMING_STOPMODE := 71,
	HOMING_TARGETPOSITION := 72,
	HOMING_VELOCITY1 := 73,
	HOMING_VELOCITY2 := 74,
	HOMING_ACCELERATION1 := 75,
	HOMING_ACCELERATION2 := 76,
	HOMING_JERK := 77,
	HOMING_TORQUELIMIT := 78,
	HOMING_TORQUETIME := 79,
	HOMING_TPCONFIG := 80,
	HOMING_RESTOREHOMEPOSITION := 81,
	HOMING_RESTORETRESHOLD := 82,
	HOMING_DRIVEHOMEMODE := 83,
	HOMING_HOMEPOSITION := 84,
	HOMING_POSSETPERMANENTLY := 85,
	HOMIN_OFFSETPOSITION := 86,
	HOMING_STOPMODEDIRECTION := 87,
	HOMESENSORDISTANCE := 88,
	CONTROLMODEDEFAULT := 90,
	ACTCONTROLMODE := 91,
	ENCODERNAME := 92,
	POSCTRLGAIN := 93,
	POSCTRLOUTPUTLIMITATION := 94,
	POSCTRKOUTPUT := 95,
	POSCTRLADAPTVALUE := 96,
	POSCTRLADAPTIONFROM0X2985 := 97,
	POSCTRLADAPTACTIVEVALUE := 98,
	SETVALUEMONITORING := 100,
	TIMELIMITSWITCHON := 101,
	REAKTONMCFBERROR := 102,
	ENABLELOGENTRY := 103,
	HWLIMITERRORREACTION := 104,
	SWLIMITERRORREACTION := 105,
	LIMITPROFILEERRORREACTION := 106,
	CINHERRORREACTION := 107,
	LIMITERSTOPREACTION := 108,
	REACTIONSSISTATUS1 := 109,
	BRAKE_MODE := 110,
	BRAKE_RELEASETIME := 111,
	BRAKE_ACTIVATIONTIME := 112,
	BRAKE_ACTMODE := 113,
	BRAKE_SAMPLEDTORQUE := 114,
	BRAKE_EFFECTIVETORQUE := 115,
	BRAKETEST_STATE := 116,
	BRAKE_SOURCESTARTVALUE := 117,
	BRAKE_MSTARTVALUE := 118,
	BRAKE_BRAKERAMPTIME := 119,
	BRAKE_BRAKEACCDEPENDING := 120,
	BRAKETEST_CMD := 121,
	BRAKETEST_MODE := 122,
	BRAKETEST_TORQUE := 123,
	BRAKETEST_THRESHOLD := 124,
	BRAKETEST_RAMPTIME := 125,
	BRAKETEST_HOLDTIME := 126,
	BRAKETEST_ACTTRESHOLD := 127,
	TORQUELIMHIGH := 128,
	TORQUELIMLOW := 129,
	WINDOWTARGETREACHED := 130,
	WINDOWTARGETREACHEDTIME := 131,
	WINDOWSTANDSTILL := 132,
	OPTIMIZEDPROFILECALCULATIONMODE := 134,
	MODPOSTOLERANCE := 135,
	RECOVERYWINDOWPOS := 136,
	RECOVERYWINDOWNEG := 137,
	SERVICEDIRECTION := 139,
	BRAKEGRINDIN_CMD := 140,
	BRAKEGRINDIN_MODE := 141,
	BRAKEGRINDIN_CTRL := 142,
	BRAKEGRINDIN_SPEED := 143,
	BRAKEGRINDIN_RAMPTIME := 144,
	BRAKEGRINDIN_ONTIME := 145,
	BRAKEGRINDIN_OFFTIME := 146,
	BRAKEGRINDIN_CYCLES := 147,
	BRAKEGRINDIN_CYCLESOUT := 148,
	BRAKEGRINDIN_STATE := 149,
	LIMITEDVELOCITY1 := 150,
	LIMITEDDECELERATION1 := 151,
	LIMITEDVELOCITY2 := 152,
	LIMITEDDECELERATION2 := 153,
	LIMITEDVELOCITY3 := 154,
	LIMITEDDECELERATION3 := 155,
	LIMITEDVELOCITY4 := 156,
	LIMITEDDECELERATION4 := 157,
	LIMITEDDISTANCE := 158,
	SLSOFFSETVELOCITY := 159,
	FOLLOWERSLS := 160,
	LIMITSPEEDCTRLSLS := 161,
	DISABLESAFETYINTERFACE := 162,
	REQUESTSAFETYINTERFACE := 163,
	SLIDISTANCE := 164,
	BRAKEGRINDIN_POSLIMIT1 := 168,
	BRAKEGRINDIN_POSLIMIT2 := 169,
	AUTOTUNING_CMD := 170,
	AT_VELOCITY := 171,
	AT_ACCELERATION := 172,
	AT_DISTANCE := 173,
	AT_CALCULATEDDISTANCE := 174,
	AT_VPNFACTOR := 175,
	AT_TNNFACTOR := 176,
	AT_STATE := 177,
	AT_VPPFACTOR := 178,
	AT_VPPFACTOREXT := 179,
	AT_WAITINGTIME := 180,
	JOGGINGSETVEL := 181,
	JOGGINGSETACC := 182,
	JOGGINGSETDEC := 183,
	JOGGINGSETJERK := 184,
	HALTDEC := 186,
	HALTJERK := 187
);
END_TYPE

(* ---- L_MC1P_PARGENERALMECHANIC.dut ---- *)
TYPE L_MC1P_PARGENERALMECHANIC :
STRUCT
	WBRAKEAVAILABLE : WORD := 0;
	LRBRAKEACTIVATIONTIME : LREAL := 0.01;
	LREXTERNALTORQUE : LREAL;
	LRBRAKEMAXTORQUE : LREAL := 2;
	LRMECHMINPOS : LREAL := 0;
	LRMECHMAXPOS : LREAL := 0;
	LRCURRCTRLPT2TT_T1 : LREAL := (246.06 * 1E-06);
	LRCURRCTRLPT2TT_T2 : LREAL := (210.35 * 1E-06);
	LRCURRCTRLPT2TT_DELAY : LREAL := (103.3 * 1E-06);
END_STRUCT
END_TYPE

(* ---- L_MC1P_PARMECHANIC.dut ---- *)
TYPE L_MC1P_PARMECHANIC :
STRUCT
	LRINERTIA : LREAL := 2.99E-05;
	LRVISCOSEFACTOR : LREAL := 0.001;
	LRCOULOMBFACTOR : LREAL := 0.025;
	LRCOULOMBSLOPE : LREAL := 1;
END_STRUCT
END_TYPE

(* ---- L_MC1P_PARMECHANIC2MS.dut ---- *)
TYPE L_MC1P_PARMECHANIC2MS :
STRUCT
	LRINERTIA2 : LREAL;
	LRD : LREAL;
	LRC : LREAL;
	LRFRICTIONRATIO : LREAL := (1.0 / 4.0);
END_STRUCT
END_TYPE

(* ---- L_MC1P_PARMECHANIC2MS_BACKLASH.dut ---- *)
TYPE L_MC1P_PARMECHANIC2MS_BACKLASH :
STRUCT
	LRBACKLASH : LREAL;
END_STRUCT
END_TYPE

(* ---- L_MC1P_PARMECHANIC3MS.dut ---- *)
TYPE L_MC1P_PARMECHANIC3MS :
STRUCT
	LRINERTIA2 : LREAL := 0.000195;
	LRINERTIA3 : LREAL := 1.6E-05;
	D1 : LREAL := 2.24;
	D2 : LREAL := 0.007;
	C1 : LREAL := 2.24;
	C2 : LREAL := 0.008;
END_STRUCT
END_TYPE

(* ---- L_MC1P_PGFUTVAL.dut ---- *)
TYPE L_MC1P_PGFUTVAL :
STRUCT
	DROUTACC : LREAL;
	DROUTSPEED : LREAL;
	DROUTPOS : LREAL;
	DRCNT : LREAL;
END_STRUCT
END_TYPE

(* ---- L_MC1P_PGPHASENPARA.dut ---- *)
TYPE L_MC1P_PGPHASENPARA :
STRUCT
	DRRELTIME : LREAL;
	DRTIME : LREAL;
	DRRELPOS : LREAL;
	DRPOS : LREAL;
	DRRELSPEED : LREAL;
	DRSPEED : LREAL;
	DRRELACC : LREAL;
	DRACC : LREAL;
	DRJERKA : LREAL;
	IBPROFILENUMBER : INT;
END_STRUCT
END_TYPE

(* ---- L_MC1P_POLEPOSITIONIDENTIFICATIONINPUT.dut ---- *)
TYPE L_MC1P_POLEPOSITIONIDENTIFICATIONINPUT :
STRUCT
	XENABLE : BOOL;
	XEXECUTEPPI : BOOL := FALSE;
	XABORTPPI : BOOL := FALSE;
	XSETPOLEPOSITION : BOOL := FALSE;
	XRESETPOLEPOSITION : BOOL := FALSE;
END_STRUCT
END_TYPE

(* ---- L_MC1P_POLEPOSITIONIDENTIFICATIONOUTPUT.dut ---- *)
TYPE L_MC1P_POLEPOSITIONIDENTIFICATIONOUTPUT :
STRUCT
	XDONE : BOOL := FALSE;
	XBUSY : BOOL := FALSE;
	XACTIVE : BOOL := FALSE;
	XCOMMANDABORTED : BOOL := FALSE;
	XERROR : BOOL := FALSE;
	EERRORID : L_IE1P_Error;
	XPPINVALID : BOOL := FALSE;
END_STRUCT
END_TYPE

(* ---- L_MC1P_POSCTRLADAPTMODE.dut ---- *)
TYPE L_MC1P_POSCTRLADAPTMODE :
(
	MOTORANDLOAD := 0,
	MOTOR := 1,
	LOAD := 2
);
END_TYPE

(* ---- L_MC1P_POSLINT.dut ---- *)
TYPE L_MC1P_POSLINT :
UNION
	LIPOS : LINT;
	ADIPOS : ARRAY [1..2] OF DINT;
END_UNION
END_TYPE

(* ---- L_MC1P_POWERINPUT.dut ---- *)
TYPE L_MC1P_POWERINPUT :
STRUCT
	ENABLE : BOOL;
	ENABLEPOSITIVE : BOOL := TRUE;
	ENABLENEGATIVE : BOOL := TRUE;
END_STRUCT
END_TYPE

(* ---- L_MC1P_POWEROUTPUT.dut ---- *)
TYPE L_MC1P_POWEROUTPUT :
STRUCT
	STATUS : BOOL;
	VALID : BOOL;
	ERROR : BOOL;
	ERRORID : L_IE1P_Error;
END_STRUCT
END_TYPE

(* ---- L_MC1P_PPISTATE.dut ---- *)
TYPE L_MC1P_PPISTATE :
(
	IDLE := 0,
	CHECKPPIACTIVATION := 1,
	PPIMONITORING := 2,
	DONE := 3,
	RESETPPIINFORMATION := 4,
	SETPPIINFORMATION := 5,
	ERROR := 999
);
END_TYPE

(* ---- L_MC1P_PRECONTROLMODE.dut ---- *)
TYPE L_MC1P_PRECONTROLMODE :
(
	AUTOMATIC := 0,
	ADDITIVEOFFSETTORQUE := 1,
	EXCLUSIVEOFFSETTORQUE := 2
);
END_TYPE

(* ---- L_MC1P_PRMDATAHEADER.dut ---- *)
TYPE L_MC1P_PRMDATAHEADER :
STRUCT
	PARAMHEADERTYPE : DWORD;
	PARAMETERDATAOFFSETFROMSTARTOF : DWORD;
	PARAMDATASIZE : DWORD;
END_STRUCT
END_TYPE

(* ---- L_MC1P_PRMFILEHEADER.dut ---- *)
TYPE L_MC1P_PRMFILEHEADER :
STRUCT
	PARSETTYPE : DWORD;
	FILEVERSION : DWORD;
	SIZETOTAL : DWORD;
	VENDOR : DWORD;
	PRODUCTCODE : DWORD;
	REVISION : DWORD;
	DATAOFFSET : DWORD;
	DATASIZE : DWORD;
	CRCCHECKSUM : DWORD;
END_STRUCT
END_TYPE

(* ---- L_MC1P_PRMPARAMETERHEADER.dut ---- *)
TYPE L_MC1P_PRMPARAMETERHEADER :
STRUCT
	SIZE : WORD;
	INDEX : WORD;
	SUBINDEX : WORD;
END_STRUCT
END_TYPE

(* ---- L_MC1P_PROFILEDATA.dut ---- *)
TYPE L_MC1P_PROFILEDATA :
STRUCT
	ALRPROFILETIME : ARRAY [0..8] OF LREAL;
	ALRPROFILEPOS : ARRAY [0..8] OF LREAL;
	ALRPROFILEVEL : ARRAY [0..8] OF LREAL;
	ALRPROFILEACC : ARRAY [0..8] OF LREAL;
	ALRPROFILEJERK : ARRAY [0..8] OF LREAL;
END_STRUCT
END_TYPE

(* ---- L_MC1P_PROFILEDATAEXTENDED.dut ---- *)
TYPE L_MC1P_PROFILEDATAEXTENDED :
STRUCT
	ALRPROFILETIME : ARRAY [0..11] OF LREAL;
	ALRPROFILEPOS : ARRAY [0..11] OF LREAL;
	ALRPROFILEVEL : ARRAY [0..11] OF LREAL;
	ALRPROFILEACC : ARRAY [0..11] OF LREAL;
	ALRPROFILEJERK : ARRAY [0..11] OF LREAL;
END_STRUCT
END_TYPE

(* ---- L_MC1P_PROFILEPARAMETER.dut ---- *)
TYPE L_MC1P_PROFILEPARAMETER :
STRUCT
	LRTARGETPOS : LREAL := 0;
	LRTARGETVEL : LREAL := 0;
	LRTARGETACC : LREAL := 0;
	LRMAXVEL : LREAL := 0;
	LRMAXACC : LREAL := 0;
	LRMAXDEC : LREAL := 0;
	LRJERKACC : LREAL := 0;
	LRJERKDEC : LREAL := 0;
END_STRUCT
END_TYPE

(* ---- L_MC1P_PROFILEPHASEDATA.dut ---- *)
TYPE L_MC1P_PROFILEPHASEDATA :
STRUCT
	T : LREAL;
	DS : LREAL;
	DV : LREAL;
	DA : LREAL;
	J : LREAL;
END_STRUCT
END_TYPE

(* ---- L_MC1P_PROFILETYPE.dut ---- *)
TYPE L_MC1P_PROFILETYPE :
(
	POLY_4TH_ORDER := 0,
	POLY_2TH_ORDER := 1,
	POLY_5TH_ORDER := 2
);
END_TYPE

(* ---- L_MC1P_QUICKSTOPOPTION.dut ---- *)
TYPE L_MC1P_QUICKSTOPOPTION :
(
	DISABLEDRIVE := 2,
	STAYINQSP := 6
);
END_TYPE

(* ---- L_MC1P_READACTUALPOSITIONINPUT.dut ---- *)
TYPE L_MC1P_READACTUALPOSITIONINPUT :
STRUCT
	ENABLE : BOOL;
END_STRUCT
END_TYPE

(* ---- L_MC1P_READACTUALPOSITIONOUTPUT.dut ---- *)
TYPE L_MC1P_READACTUALPOSITIONOUTPUT :
STRUCT
	VALID : BOOL;
	BUSY : BOOL;
	ERROR : BOOL;
	ERRORID : L_IE1P_Error;
	POSITION : LREAL;
END_STRUCT
END_TYPE

(* ---- L_MC1P_READACTUALTORQUEINPUT.dut ---- *)
TYPE L_MC1P_READACTUALTORQUEINPUT :
STRUCT
	ENABLE : BOOL;
END_STRUCT
END_TYPE

(* ---- L_MC1P_READACTUALTORQUEOUTPUT.dut ---- *)
TYPE L_MC1P_READACTUALTORQUEOUTPUT :
STRUCT
	VALID : BOOL;
	BUSY : BOOL;
	ERROR : BOOL;
	ERRORID : L_IE1P_Error;
	TORQUE : LREAL;
END_STRUCT
END_TYPE

(* ---- L_MC1P_READACTUALVELOCITYINPUT.dut ---- *)
TYPE L_MC1P_READACTUALVELOCITYINPUT :
STRUCT
	ENABLE : BOOL;
END_STRUCT
END_TYPE

(* ---- L_MC1P_READACTUALVELOCITYOUTPUT.dut ---- *)
TYPE L_MC1P_READACTUALVELOCITYOUTPUT :
STRUCT
	VALID : BOOL;
	BUSY : BOOL;
	ERROR : BOOL;
	ERRORID : L_IE1P_Error;
	VELOCITY : LREAL;
END_STRUCT
END_TYPE

(* ---- L_MC1P_READAXISERRORINPUT.dut ---- *)
TYPE L_MC1P_READAXISERRORINPUT :
STRUCT
	ENABLE : BOOL;
END_STRUCT
END_TYPE

(* ---- L_MC1P_READAXISERROROUTPUT.dut ---- *)
TYPE L_MC1P_READAXISERROROUTPUT :
STRUCT
	VALID : BOOL;
	BUSY : BOOL;
	ERROR : BOOL;
	ERRORID : L_IE1P_Error;
	AXISWARNING : BOOL;
	AXISERROR : BOOL;
	AXISERRORID : L_IE1P_Error;
	PINSTANCENAME : POINTER TO STRING;
	TIMESTAMP : TIME;
	DRIVEWARNING : BOOL;
	DRIVEERROR : BOOL;
	DRIVEERRORID : DWORD;
END_STRUCT
END_TYPE

(* ---- L_MC1P_READAXISINFOINPUT.dut ---- *)
TYPE L_MC1P_READAXISINFOINPUT :
STRUCT
	ENABLE : BOOL;
END_STRUCT
END_TYPE

(* ---- L_MC1P_READAXISINFOOUTPUT.dut ---- *)
TYPE L_MC1P_READAXISINFOOUTPUT :
STRUCT
	VALID : BOOL;
	BUSY : BOOL;
	ERROR : BOOL;
	ERRORID : L_IE1P_Error;
	HOMEABSSWITCH : BOOL;
	LIMITSWITCHPOS : BOOL;
	LIMITSWITCHNEG : BOOL;
	SIMULATION : BOOL;
	COMMUNICATIONREADY : BOOL;
	READYFORPOWERON : BOOL;
	POWERON : BOOL;
	ISHOMED : BOOL;
	AXISERROR : BOOL;
	AXISWARNING : BOOL;
	DRIVEWARNING : BOOL;
	DRIVEERROR : BOOL;
	SWLIMITSWITCHPOS : BOOL;
	SWLIMITSWITCHNEG : BOOL;
	READYFORMOTION : BOOL;
	STOACTIVE : BOOL;
	VOLTAGEENABLED : BOOL;
	MOTORMAGNETISED : BOOL;
	QSPAPPLACTIVE : BOOL;
	QSPDRIVEACTIVE : BOOL;
END_STRUCT
END_TYPE

(* ---- L_MC1P_READAXISSTATUSWORDSINPUT.dut ---- *)
TYPE L_MC1P_READAXISSTATUSWORDSINPUT :
STRUCT
	XENABLE : BOOL;
END_STRUCT
END_TYPE

(* ---- L_MC1P_READAXISSTATUSWORDSOUTPUT.dut ---- *)
TYPE L_MC1P_READAXISSTATUSWORDSOUTPUT :
STRUCT
	XVALID : BOOL;
	XBUSY : BOOL;
	XERROR : BOOL;
	EERRORID : L_IE1P_Error;
	WCIA402STATUSWORD : WORD;
	WLENZESTATUSWORD : WORD;
	WLENZESTATUSWORD2 : WORD;
	WLENZESTATUSWORDEXT : WORD;
END_STRUCT
END_TYPE

(* ---- L_MC1P_READBOOLPARAMETERINPUT.dut ---- *)
TYPE L_MC1P_READBOOLPARAMETERINPUT :
STRUCT
	ENABLE : BOOL;
	PARAMETERNUMBER : DINT;
	TCYCLETIME : TIME;
END_STRUCT
END_TYPE

(* ---- L_MC1P_READBOOLPARAMETEROUTPUT.dut ---- *)
TYPE L_MC1P_READBOOLPARAMETEROUTPUT :
STRUCT
	VALID : BOOL;
	BUSY : BOOL;
	ERROR : BOOL;
	ERRORID : L_IE1P_Error;
	VALUE : BOOL;
END_STRUCT
END_TYPE

(* ---- L_MC1P_READMACHINEDATAINPUT.dut ---- *)
TYPE L_MC1P_READMACHINEDATAINPUT :
STRUCT
	XENABLE : BOOL;
END_STRUCT
END_TYPE

(* ---- L_MC1P_READMACHINEDATAOUTPUT.dut ---- *)
TYPE L_MC1P_READMACHINEDATAOUTPUT :
STRUCT
	XVALID : BOOL;
	XBUSY : BOOL;
	XERROR : BOOL;
	EERRORID : L_IE1P_Error;
	LRFEEDCONSTANT : LREAL;
	DWGEARDENOMINATOR : DWORD;
	DWGEARNUMERATOR : DWORD;
	DWADDGEARDENOMINATOR : DWORD;
	DWADDGEARNUMERATOR : DWORD;
	DWPOSRESOLUTION : DWORD;
	XORIENTATION : BOOL;
	ETRAVERSINGRANGE : L_MC1P_TraversingRange;
	LRCYCLELENGTH : LREAL;
	XVIRTUAL : BOOL;
END_STRUCT
END_TYPE

(* ---- L_MC1P_READMOTIONSTATEINPUT.dut ---- *)
TYPE L_MC1P_READMOTIONSTATEINPUT :
STRUCT
	ENABLE : BOOL;
	SOURCE : MC_SOURCE;
END_STRUCT
END_TYPE

(* ---- L_MC1P_READMOTIONSTATEOUTPUT.dut ---- *)
TYPE L_MC1P_READMOTIONSTATEOUTPUT :
STRUCT
	VALID : BOOL;
	BUSY : BOOL;
	ERROR : BOOL;
	ERRORID : L_IE1P_Error;
	CONSTANTVELOCITY : BOOL;
	ACCELERATING : BOOL;
	DECELERATING : BOOL;
	DIRECTIONPOSITIVE : BOOL;
	DIRECTIONNEGATIVE : BOOL;
	INPOSITION : BOOL;
	STANDSTILLSETVELOCITY : BOOL;
	STANDSTILLACTVELOCITY : BOOL;
END_STRUCT
END_TYPE

(* ---- L_MC1P_READPARAMETERINPUT.dut ---- *)
TYPE L_MC1P_READPARAMETERINPUT :
STRUCT
	ENABLE : BOOL;
	PARAMETERNUMBER : DINT;
	TCYCLETIME : TIME := TIME#1ms;
END_STRUCT
END_TYPE

(* ---- L_MC1P_READPARAMETEROUTPUT.dut ---- *)
TYPE L_MC1P_READPARAMETEROUTPUT :
STRUCT
	VALID : BOOL;
	BUSY : BOOL;
	ERROR : BOOL;
	ERRORID : L_IE1P_Error;
	VALUE : LREAL;
END_STRUCT
END_TYPE

(* ---- L_MC1P_READSETPOSITIONINPUT.dut ---- *)
TYPE L_MC1P_READSETPOSITIONINPUT :
STRUCT
	XENABLE : BOOL;
END_STRUCT
END_TYPE

(* ---- L_MC1P_READSETPOSITIONOUTPUT.dut ---- *)
TYPE L_MC1P_READSETPOSITIONOUTPUT :
STRUCT
	XVALID : BOOL;
	XBUSY : BOOL;
	XERROR : BOOL;
	EERRORID : L_IE1P_Error;
	LRPOSITION : LREAL;
END_STRUCT
END_TYPE

(* ---- L_MC1P_READSTATUSINPUT.dut ---- *)
TYPE L_MC1P_READSTATUSINPUT :
STRUCT
	ENABLE : BOOL;
END_STRUCT
END_TYPE

(* ---- L_MC1P_READSTATUSOUTPUT.dut ---- *)
TYPE L_MC1P_READSTATUSOUTPUT :
STRUCT
	VALID : BOOL;
	BUSY : BOOL;
	ERROR : BOOL;
	ERRORID : L_IE1P_Error;
	ERRORSTOP : BOOL;
	DISABLED : BOOL;
	STOPPING : BOOL;
	HOMING : BOOL;
	STANDSTILL : BOOL;
	DISCRETEMOTION : BOOL;
	CONTINUOUSMOTION : BOOL;
	SYNCHRONIZEDMOTION : BOOL;
	CONSTANTVELOCITY : BOOL;
	ACCELERATING : BOOL;
	DECELERATING : BOOL;
	INPOSITION : BOOL;
END_STRUCT
END_TYPE

(* ---- L_MC1P_REINITNODEINPUT.dut ---- *)
TYPE L_MC1P_REINITNODEINPUT :
STRUCT
	XEXECUTE : BOOL;
END_STRUCT
END_TYPE

(* ---- L_MC1P_REINITNODEOUTPUT.dut ---- *)
TYPE L_MC1P_REINITNODEOUTPUT :
STRUCT
	XDONE : BOOL;
	XBUSY : BOOL;
	XERROR : BOOL;
	EERRORID : L_IE1P_Error;
END_STRUCT
END_TYPE

(* ---- L_MC1P_RESETFOLLOWINGERRORINPUT.dut ---- *)
TYPE L_MC1P_RESETFOLLOWINGERRORINPUT :
STRUCT
	XEXECUTE : BOOL;
END_STRUCT
END_TYPE

(* ---- L_MC1P_RESETFOLLOWINGERROROUTPUT.dut ---- *)
TYPE L_MC1P_RESETFOLLOWINGERROROUTPUT :
STRUCT
	XDONE : BOOL;
	XERROR : BOOL;
	EERRORID : L_IE1P_Error;
END_STRUCT
END_TYPE

(* ---- L_MC1P_RESETHOMEPOSITIONINPUT.dut ---- *)
TYPE L_MC1P_RESETHOMEPOSITIONINPUT :
STRUCT
	XEXECUTE : BOOL;
	XRESETPOSITIONOFFSET : BOOL;
END_STRUCT
END_TYPE

(* ---- L_MC1P_RESETHOMEPOSITIONOUTPUT.dut ---- *)
TYPE L_MC1P_RESETHOMEPOSITIONOUTPUT :
STRUCT
	XDONE : BOOL;
	XBUSY : BOOL;
	XERROR : BOOL;
	EERRORID : L_IE1P_Error;
END_STRUCT
END_TYPE

(* ---- L_MC1P_RESETINPUT.dut ---- *)
TYPE L_MC1P_RESETINPUT :
STRUCT
	EXECUTE : BOOL;
END_STRUCT
END_TYPE

(* ---- L_MC1P_RESETOUTPUT.dut ---- *)
TYPE L_MC1P_RESETOUTPUT :
STRUCT
	DONE : BOOL;
	BUSY : BOOL;
	ERROR : BOOL;
	ERRORID : L_IE1P_Error;
END_STRUCT
END_TYPE

(* ---- L_MC1P_RETAINDATAENCAXIS.dut ---- *)
TYPE L_MC1P_RETAINDATAENCAXIS :
STRUCT
	XRETAININITIALIZED : BOOL;
	RETAINSTACK1 : L_MC1P_uRetainData;
	RETAINSTACK2 : L_MC1P_uRetainData;
END_STRUCT
END_TYPE

(* ---- L_MC1P_RETAINDATAI700.dut ---- *)
TYPE L_MC1P_RETAINDATAI700 :
STRUCT
	DWENCODERCRC : DWORD;
	LRBRAKESAMPLEDTORQUE : LREAL;
END_STRUCT
END_TYPE

(* ---- L_MC1P_RETAINDATAI700_V2.dut ---- *)
TYPE L_MC1P_RETAINDATAI700_V2 :
STRUCT
	DWENCODERCRC : DWORD;
	LRBRAKESAMPLEDTORQUE : LREAL;
END_STRUCT
END_TYPE

(* ---- L_MC1P_RETAINDATAI700_V3.dut ---- *)
TYPE L_MC1P_RETAINDATAI700_V3 :
STRUCT
	DWENCODERCRC : DWORD;
	LRBRAKESAMPLEDTORQUE : LREAL;
END_STRUCT
END_TYPE

(* ---- L_MC1P_RETAINDATAREALDRIVE.dut ---- *)
TYPE L_MC1P_RETAINDATAREALDRIVE :
STRUCT
	DWPROPERTIES : DWORD;
	UPOSACT : L_MC1P_PosLINT;
	DIREFOFFSETINC : DINT;
	LRACTPOS : LREAL;
	LRABSREFOFFSET : LREAL;
	LRCYCLELENGTH : LREAL;
	LRSCALEFACTOR : LREAL;
END_STRUCT
END_TYPE

(* ---- L_MC1P_RETAINDATAREALDRIVE_V2.dut ---- *)
TYPE L_MC1P_RETAINDATAREALDRIVE_V2 :
STRUCT
	DWPROPERTIES : DWORD;
	UPOSACT : L_MC1P_PosLINT;
	DIREFOFFSETINC : DINT;
	LRACTPOS : LREAL;
	LRABSREFOFFSET : LREAL;
	LRCYCLELENGTH : LREAL;
	LRSCALEFACTOR : LREAL;
	DISETPOSROUNDSLAST : DINT;
	LRLASTSETPOSITION : LREAL;
	DITARGETPOSROUNDS : DINT;
	LRLASTTARGETPOSITION : LREAL;
END_STRUCT
END_TYPE

(* ---- L_MC1P_RETAINDATAREALDRIVE_V3.dut ---- *)
TYPE L_MC1P_RETAINDATAREALDRIVE_V3 :
STRUCT
	DWPROPERTIES : DWORD;
	DIREFOFFSETINC : DINT;
	UPOSACT : L_MC1P_PosLINT;
	LRACTPOS : LREAL;
	LRABSREFOFFSET : LREAL;
	LRCYCLELENGTH : LREAL;
	LRSCALEFACTOR : LREAL;
	LRLASTSETPOSITION : LREAL;
	DISETPOSROUNDSLAST : DINT;
	DITARGETPOSROUNDS : DINT;
	LRLASTTARGETPOSITION : LREAL;
	DRIVEGUID : L_MC1P_AxisGUID;
END_STRUCT
END_TYPE

(* ---- L_MC1P_RETAINDATATYPE.dut ---- *)
TYPE L_MC1P_RETAINDATATYPE :
(
	NONE := -1,
	DATAREALDRIVE := 0,
	DATAI700 := 1
);
END_TYPE

(* ---- L_MC1P_SAFETYREADSTATUSWORDSINPUT.dut ---- *)
TYPE L_MC1P_SAFETYREADSTATUSWORDSINPUT :
STRUCT
	XENABLE : BOOL;
END_STRUCT
END_TYPE

(* ---- L_MC1P_SAFETYREADSTATUSWORDSOUTPUT.dut ---- *)
TYPE L_MC1P_SAFETYREADSTATUSWORDSOUTPUT :
STRUCT
	XVALID : BOOL;
	XBUSY : BOOL;
	XERROR : BOOL;
	EERRORID : L_IE1P_Error;
	DWCONTROL : DWORD;
	DWSTATE : DWORD;
	DWIOSTATE : DWORD;
END_STRUCT
END_TYPE

(* ---- L_MC1P_SCALEFIXTOLREAL.dut ---- *)
TYPE L_MC1P_SCALEFIXTOLREAL :
(
	NONE := 0,
	FIX_X := 1,
	FIX_X_X := 10,
	FIX_X_XX := 100,
	FIX_X_XXX := 1000,
	FIX_X_XXXX := 10000,
	FIX_X_XXXXX := 100000
);
END_TYPE

(* ---- L_MC1P_SERVICEDIRECTION.dut ---- *)
TYPE L_MC1P_SERVICEDIRECTION :
(
	BOTH := 0,
	POSITIVE := 1,
	NEGATIVE := 2
);
END_TYPE

(* ---- L_MC1P_SETBASICPARAMETERINPUT.dut ---- *)
TYPE L_MC1P_SETBASICPARAMETERINPUT :
STRUCT
	XENABLE : BOOL;
	XSETJOGPARAMETER : BOOL;
	LRJOGVEL : LREAL := 360;
	LRJOGACC : LREAL := 360;
	LRJOGDEC : LREAL := 1440;
	LRJOGJERK : LREAL := 0;
	XSETHALTPARAMETER : BOOL;
	LRHALTDEC : LREAL := 1800;
	LRHALTJERK : LREAL := 0;
	XSETQSPAPPLPARAMETER : BOOL;
	LRQSPAPPLDEC : LREAL := 3600.0;
	LRQSPAPPLJERK : LREAL := 0;
	XSETHOMEPOSITION : BOOL;
	LRHOMEPOSITION : LREAL;
	XSETHOMEPARAMETER : BOOL;
	SCHOMEPARAMETER : L_MC1P_HomeParameter := STRUCT(eHomeMode := L_MC1P_HomeMode.SetPositionDirect, eHomeStopMode := L_MC1P_HomeStopMode.StopPositioning, lrTargetPosition := 0, lrVelocity1 := 360.0, lrVelocity2 := 0, lrAcceleration1 := 720.0, lrAcceleration2 := 360.0, lrJerk := 7200.0, rTorqueLimit := 0.1, rTorqueTime := 1.0, dwTPConfig := 1, eStopModeDirection := MC_DIRECTION.mcCurrentDirection);
END_STRUCT
END_TYPE

(* ---- L_MC1P_SETBASICPARAMETEROUTPUT.dut ---- *)
TYPE L_MC1P_SETBASICPARAMETEROUTPUT :
STRUCT
	XBUSY : BOOL;
	XERROR : BOOL;
	EERRORID : L_IE1P_Error;
END_STRUCT
END_TYPE

(* ---- L_MC1P_SETCONTROLMODEINPUT.dut ---- *)
TYPE L_MC1P_SETCONTROLMODEINPUT :
STRUCT
	XEXECUTE : BOOL;
	ECONTROLMODE : L_MC1P_ControlModeSet := L_MC1P_ControlModeSet.PosCtrlDrive;
	XKEEPACTPOSPRIORFDB : BOOL := FALSE;
	XRESTARTPOSITIONING : BOOL := FALSE;
END_STRUCT
END_TYPE

(* ---- L_MC1P_SETCONTROLMODEOUTPUT.dut ---- *)
TYPE L_MC1P_SETCONTROLMODEOUTPUT :
STRUCT
	XDONE : BOOL;
	XBUSY : BOOL;
	XERROR : BOOL;
	EERRORID : L_IE1P_Error;
END_STRUCT
END_TYPE

(* ---- L_MC1P_SETDCBRAKEINPUT.dut ---- *)
TYPE L_MC1P_SETDCBRAKEINPUT :
STRUCT
	XENABLE : BOOL;
END_STRUCT
END_TYPE

(* ---- L_MC1P_SETDCBRAKEOUTPUT.dut ---- *)
TYPE L_MC1P_SETDCBRAKEOUTPUT :
STRUCT
	XBUSY : BOOL;
	XACTIVE : BOOL;
	XERROR : BOOL;
	EERRORID : L_IE1P_Error;
END_STRUCT
END_TYPE

(* ---- L_MC1P_SETINERTIAADAPTVALUEINPUT.dut ---- *)
TYPE L_MC1P_SETINERTIAADAPTVALUEINPUT :
STRUCT
	XENABLE : BOOL;
	LRINERTIAADAPTVALUE : LREAL := 1.0;
END_STRUCT
END_TYPE

(* ---- L_MC1P_SETINERTIAADAPTVALUEOUTPUT.dut ---- *)
TYPE L_MC1P_SETINERTIAADAPTVALUEOUTPUT :
STRUCT
	XBUSY : BOOL;
	XERROR : BOOL;
	EERRORID : L_IE1P_Error;
END_STRUCT
END_TYPE

(* ---- L_MC1P_SETOVERRIDEINPUT.dut ---- *)
TYPE L_MC1P_SETOVERRIDEINPUT :
STRUCT
	ENABLE : BOOL;
	VELFACTOR : LREAL := 1.0;
	ACCFACTOR : LREAL := 1.0;
	JERKFACTOR : LREAL := 1.0;
END_STRUCT
END_TYPE

(* ---- L_MC1P_SETOVERRIDEOUTPUT.dut ---- *)
TYPE L_MC1P_SETOVERRIDEOUTPUT :
STRUCT
	ENABLED : BOOL;
	BUSY : BOOL;
	ERROR : BOOL;
	ERRORID : L_IE1P_Error;
END_STRUCT
END_TYPE

(* ---- L_MC1P_SETPOSCTRLADAPTVALUEINPUT.dut ---- *)
TYPE L_MC1P_SETPOSCTRLADAPTVALUEINPUT :
STRUCT
	XENABLE : BOOL;
	LRPOSCTRLADAPTVALUE : LREAL := 1.0;
	EMODE : L_MC1P_PosCtrlAdaptMode := L_MC1P_PosCtrlAdaptMode.MotorAndLoad;
END_STRUCT
END_TYPE

(* ---- L_MC1P_SETPOSCTRLADAPTVALUEOUTPUT.dut ---- *)
TYPE L_MC1P_SETPOSCTRLADAPTVALUEOUTPUT :
STRUCT
	XBUSY : BOOL;
	XERROR : BOOL;
	EERRORID : L_IE1P_Error;
END_STRUCT
END_TYPE

(* ---- L_MC1P_SETPOSITIONINPUT.dut ---- *)
TYPE L_MC1P_SETPOSITIONINPUT :
STRUCT
	EXECUTE : BOOL;
	POSITION : LREAL;
	RELATIVE : BOOL;
	EXECUTIONMODE : MC_EXECUTION_MODE := MC_EXECUTION_MODE.mcImmediately;
	RESTARTPOSITIONING : BOOL := FALSE;
	USESETTINGSFROMHOMINGMODE : BOOL := FALSE;
	XCALLFROMAXESGROUP : BOOL;
	XDISABLELOGMESSAGE : BOOL;
END_STRUCT
END_TYPE

(* ---- L_MC1P_SETPOSITIONOUTPUT.dut ---- *)
TYPE L_MC1P_SETPOSITIONOUTPUT :
STRUCT
	DONE : BOOL;
	BUSY : BOOL;
	ERROR : BOOL;
	ERRORID : L_IE1P_Error;
END_STRUCT
END_TYPE

(* ---- L_MC1P_SETQUICKSTOPAPPLINPUT.dut ---- *)
TYPE L_MC1P_SETQUICKSTOPAPPLINPUT :
STRUCT
	XENABLE : BOOL;
END_STRUCT
END_TYPE

(* ---- L_MC1P_SETQUICKSTOPAPPLOUTPUT.dut ---- *)
TYPE L_MC1P_SETQUICKSTOPAPPLOUTPUT :
STRUCT
	XBUSY : BOOL;
	XACTIVE : BOOL;
	XERROR : BOOL;
	EERRORID : L_IE1P_Error;
END_STRUCT
END_TYPE

(* ---- L_MC1P_SETQUICKSTOPINPUT.dut ---- *)
TYPE L_MC1P_SETQUICKSTOPINPUT :
STRUCT
	XENABLE : BOOL;
END_STRUCT
END_TYPE

(* ---- L_MC1P_SETQUICKSTOPOPTIONINPUT.dut ---- *)
TYPE L_MC1P_SETQUICKSTOPOPTIONINPUT :
STRUCT
	XEXECUTE : BOOL;
	EQUICKSTOPOPTION : L_MC1P_QuickStopOption := L_MC1P_QuickStopOption.StayInQSP;
END_STRUCT
END_TYPE

(* ---- L_MC1P_SETQUICKSTOPOPTIONOUTPUT.dut ---- *)
TYPE L_MC1P_SETQUICKSTOPOPTIONOUTPUT :
STRUCT
	XDONE : BOOL;
	XBUSY : BOOL;
	XERROR : BOOL;
	EERRORID : L_IE1P_Error;
END_STRUCT
END_TYPE

(* ---- L_MC1P_SETQUICKSTOPOUTPUT.dut ---- *)
TYPE L_MC1P_SETQUICKSTOPOUTPUT :
STRUCT
	XBUSY : BOOL;
	XACTIVE : BOOL;
	XERROR : BOOL;
	EERRORID : L_IE1P_Error;
END_STRUCT
END_TYPE

(* ---- L_MC1P_SETSPEEDCTRLADAPTVALUEINPUT.dut ---- *)
TYPE L_MC1P_SETSPEEDCTRLADAPTVALUEINPUT :
STRUCT
	XENABLE : BOOL;
	LRSPEEDCTRLADAPTVALUE : LREAL := 1.0;
END_STRUCT
END_TYPE

(* ---- L_MC1P_SETSPEEDCTRLADAPTVALUEOUTPUT.dut ---- *)
TYPE L_MC1P_SETSPEEDCTRLADAPTVALUEOUTPUT :
STRUCT
	XBUSY : BOOL;
	XERROR : BOOL;
	EERRORID : L_IE1P_Error;
END_STRUCT
END_TYPE

(* ---- L_MC1P_SETSPEEDCTRLLOADVALUEINPUT.dut ---- *)
TYPE L_MC1P_SETSPEEDCTRLLOADVALUEINPUT :
STRUCT
	XENABLE : BOOL;
	LRSPEEDCTRLLOADVALUE : LREAL := 1.0;
END_STRUCT
END_TYPE

(* ---- L_MC1P_SETSPEEDCTRLLOADVALUEOUTPUT.dut ---- *)
TYPE L_MC1P_SETSPEEDCTRLLOADVALUEOUTPUT :
STRUCT
	XBUSY : BOOL;
	XERROR : BOOL;
	EERRORID : L_IE1P_Error;
END_STRUCT
END_TYPE

(* ---- L_MC1P_SETTORQUELIMITINPUT.dut ---- *)
TYPE L_MC1P_SETTORQUELIMITINPUT :
STRUCT
	XENABLE : BOOL;
	XSETTORQUELIMITPOS : BOOL;
	LRTORQUELIMITPOS : LREAL;
	XSETTORQUELIMITNEG : BOOL;
	LRTORQUELIMITNEG : LREAL;
	XTORQUEINPUTASPERCENT : BOOL;
END_STRUCT
END_TYPE

(* ---- L_MC1P_SETTORQUELIMITOUTPUT.dut ---- *)
TYPE L_MC1P_SETTORQUELIMITOUTPUT :
STRUCT
	XBUSY : BOOL;
	XERROR : BOOL;
	EERRORID : L_IE1P_Error;
END_STRUCT
END_TYPE

(* ---- L_MC1P_SETTORQUEOFFSETINPUT.dut ---- *)
TYPE L_MC1P_SETTORQUEOFFSETINPUT :
STRUCT
	XENABLE : BOOL;
	LRTORQUE : LREAL;
	EPRECONTROLMODE : L_MC1P_PreControlMode := L_MC1P_PreControlMode.AdditiveOffsetTorque;
END_STRUCT
END_TYPE

(* ---- L_MC1P_SETTORQUEOFFSETOUTPUT.dut ---- *)
TYPE L_MC1P_SETTORQUEOFFSETOUTPUT :
STRUCT
	XBUSY : BOOL;
	XERROR : BOOL;
	EERRORID : L_IE1P_Error;
END_STRUCT
END_TYPE

(* ---- L_MC1P_SETVALUEMODE.dut ---- *)
TYPE L_MC1P_SETVALUEMODE :
(
	POS := 1,
	VEL := 2,
	POSVEL := 3,
	VELACC := 6,
	POSVELACC := 7,
	VEL_VELFROMPROFILEGEN := 8,
	VEL_VELFROMDIFFPOS := 9,
	POSDIFFVELACC := 10
);
END_TYPE

(* ---- L_MC1P_SIMAXISCYCLETIME.dut ---- *)
TYPE L_MC1P_SIMAXISCYCLETIME :
(
	TASKCYCLE_1KHZ := 1,
	TASKCYCLE_2KHZ := 2,
	TASKCYCLE_4KHZ := 4,
	TASKCYCLE_8KHZ := 8,
	TASKCYCLE_16KHZ := 16,
	TASKCYCLE_32KHZ := 32,
	TASKCYCLE_64KHZ := 64
);
END_TYPE

(* ---- L_MC1P_STATUSABC.dut ---- *)
TYPE L_MC1P_STATUSABC :
STRUCT
	XINTERNALCONTROLACTIVE : BOOL;
	XERROR : BOOL;
	EERRORID : L_IE1P_Error;
	XFUNBUSY : BOOL;
	XFUNDONE : BOOL;
	XFUNCOMMANDABORTED : BOOL;
	EFUNSTATEACT : L_MC1P_ABC_State;
	ECONTROLMODE : L_MC1P_ControlMode;
	XISHOMED : BOOL;
	XHWLIMITSWITCHNEG : BOOL;
	XHWLIMITSWITCHPOS : BOOL;
	XSWLIMITENABLED : BOOL;
	XSWLIMITSWITCHNEG : BOOL;
	XSWLIMITSWITCHPOS : BOOL;
	EAXISTYPE : L_MC1P_DriveType;
	EAXISSTATE : L_MC1P_AXIS_STATE;
	XAXISREADY : BOOL;
	XAXISENABLED : BOOL;
	XAXISWARNING : BOOL;
	XAXISERROR : BOOL;
	EAXISERRORID : L_IE1P_Error;
	XDRIVEWARNING : BOOL;
	XDRIVEERROR : BOOL;
	DWDRIVEERRORID : DWORD;
	LRACTPOS : LREAL;
	LRACTVEL : LREAL;
	LRSETPOSOUT : LREAL;
	LRSETVELOUT : LREAL;
	LRACTFOLLOWINGERROR : LREAL;
	XCONSTANTVELOCITY : BOOL;
	XACCELERATING : BOOL;
	XDECELERATING : BOOL;
	XDIRECTIONPOSITIVE : BOOL;
	XDIRECTIONNEGATIVE : BOOL;
	XINPOSITION : BOOL;
	XAXISAVAILABLE : BOOL;
	XSTANDSTILLSETVELOCITY : BOOL;
	XSTANDSTILLACTVELOCITY : BOOL;
	XAXISREADYTOSWITCHON : BOOL;
	XAXISREADYFORMOTION : BOOL;
END_STRUCT
END_TYPE

(* ---- L_MC1P_STATUSAXIS.dut ---- *)
TYPE L_MC1P_STATUSAXIS :
STRUCT
	XJOGACTIVE : BOOL;
	ECONTROLMODE : L_MC1P_ControlMode := L_MC1P_ControlMode.PosCtrlDrive;
	XISHOMED : BOOL;
	XHWLIMITSWITCHNEG : BOOL;
	XHWLIMITSWITCHPOS : BOOL;
	XSWLIMITENABLED : BOOL;
	XSWLIMITSWITCHNEG : BOOL;
	XSWLIMITSWITCHPOS : BOOL;
	EAXISTYPE : L_MC1P_DriveType := L_MC1P_DriveType.Virtual;
	EAXISSTATE : L_MC1P_AXIS_STATE := L_MC1P_AXIS_STATE.Disabled;
	XSTOACTIVE : BOOL;
	XREADYFOROPERATION : BOOL;
	XOPERATIONENABLED : BOOL;
	XREADYFORMOTION : BOOL;
	XAXISWARNING : BOOL;
	XAXISERROR : BOOL;
	EAXISERRORID : L_IE1P_Error;
	XDRIVEWARNING : BOOL;
	XDRIVEERROR : BOOL;
	DWDRIVEERRORID : DWORD;
	LRACTPOS : LREAL;
	LRACTVEL : LREAL;
	LRSETPOSOUT : LREAL;
	LRSETVELOUT : LREAL;
	LRACTFOLLOWINGERROR : LREAL;
	XINPOSITION : BOOL;
	XSTANDSTILLSETVELOCITY : BOOL;
	XSTANDSTILLACTVELOCITY : BOOL;
	XCONSTANTVELOCITY : BOOL;
	XACCELERATING : BOOL;
	XDECELERATING : BOOL;
	XDIRECTIONPOSITIVE : BOOL;
	XDIRECTIONNEGATIVE : BOOL;
	XAXISAVAILABLE : BOOL;
END_STRUCT
END_TYPE

(* ---- L_MC1P_STOPINPUT.dut ---- *)
TYPE L_MC1P_STOPINPUT :
STRUCT
	EXECUTE : BOOL;
	DECELERATION : LREAL;
	JERK : LREAL;
END_STRUCT
END_TYPE

(* ---- L_MC1P_STOPOPERATION.dut ---- *)
TYPE L_MC1P_STOPOPERATION :
STRUCT
	XSETQSP : BOOL;
	XSETQSPCINH : BOOL;
	XSETCINH : BOOL;
	XSETFASTSTOP : BOOL;
END_STRUCT
END_TYPE

(* ---- L_MC1P_STOPOUTPUT.dut ---- *)
TYPE L_MC1P_STOPOUTPUT :
STRUCT
	DONE : BOOL;
	BUSY : BOOL;
	COMMANDABORTED : BOOL;
	ERROR : BOOL;
	ERRORID : L_IE1P_Error;
	XUSED : BOOL;
END_STRUCT
END_TYPE

(* ---- L_MC1P_SUSPENDFOLLOWINGERRORINPUT.dut ---- *)
TYPE L_MC1P_SUSPENDFOLLOWINGERRORINPUT :
STRUCT
	XENABLE : BOOL;
END_STRUCT
END_TYPE

(* ---- L_MC1P_SUSPENDFOLLOWINGERROROUTPUT.dut ---- *)
TYPE L_MC1P_SUSPENDFOLLOWINGERROROUTPUT :
STRUCT
	XBUSY : BOOL;
	XERROR : BOOL;
	EERRORID : L_IE1P_Error;
END_STRUCT
END_TYPE

(* ---- L_MC1P_TEMPLATE_EDGEINPUT.dut ---- *)
TYPE L_MC1P_TEMPLATE_EDGEINPUT :
STRUCT
	XEXECUTE : BOOL;
END_STRUCT
END_TYPE

(* ---- L_MC1P_TEMPLATE_EDGEOUTPUT.dut ---- *)
TYPE L_MC1P_TEMPLATE_EDGEOUTPUT :
STRUCT
	XDONE : BOOL;
	XBUSY : BOOL;
	XCOMMANDABORTED : BOOL;
	XERROR : BOOL;
	EERRORID : L_IE1P_Error;
END_STRUCT
END_TYPE

(* ---- L_MC1P_TIMESTAMP.dut ---- *)
TYPE L_MC1P_TIMESTAMP :
STRUCT
	TIME_01 : SysTime;
	TIME_02 : SysTime;
	TIME_03 : SysTime;
	TIME_04 : SysTime;
	TIME_05 : SysTime;
	TIME_06 : SysTime;
	TIME_07 : SysTime;
	TIME_08 : SysTime;
	TIME_DELTA_01_02 : SysTime;
	TIME_DELTA_02_03 : SysTime;
	TIME_DELTA_03_04 : SysTime;
	TIME_DELTA_04_05 : SysTime;
	TIME_DELTA_05_06 : SysTime;
	TIME_DELTA_06_07 : SysTime;
	TIME_DELTA_07_08 : SysTime;
END_STRUCT
END_TYPE

(* ---- L_MC1P_TORQUECONTROLINPUT.dut ---- *)
TYPE L_MC1P_TORQUECONTROLINPUT :
STRUCT
	XCONTINUOUSUPDATE : BOOL := TRUE;
	LRTORQUE : LREAL := 0;
	LRVELOCITYLIMITHIGH : LREAL := 0;
	LRVELOCITYLIMITLOW : LREAL := 0;
	XVALIDATESPEEDLIMITS : BOOL := TRUE;
END_STRUCT
END_TYPE

(* ---- L_MC1P_TORQUECONTROLOUTPUT.dut ---- *)
TYPE L_MC1P_TORQUECONTROLOUTPUT :
STRUCT
END_STRUCT
END_TYPE

(* ---- L_MC1P_TORQUETESTMONITORING.dut ---- *)
TYPE L_MC1P_TORQUETESTMONITORING :
STRUCT
	PT1_ACTMOTORTORQUE : L_USPP_PT1Filter;
	PT1_SETTORQUE : L_USPP_PT1Filter;
	LRPT1DELAY : LREAL := 0.01;
	ALRSETTORQUE : ARRAY [0..15] OF LREAL;
	LRTORQUETOLERANCE : LREAL := 0.1;
	IDX : UINT;
	XBUFFER : BOOL;
END_STRUCT
END_TYPE

(* ---- L_MC1P_TORQUETESTSEQUENCE.dut ---- *)
TYPE L_MC1P_TORQUETESTSEQUENCE :
(
	ETT_DEFAULT := 0,
	ETT_PREINIT := 9,
	ETT_INIT := 1,
	ETT_CONTROLMODE := 2,
	ETT_TORQUERAMPUP := 3,
	ETT_TORQUERAMPDOWN := 4,
	ETT_CONSTANTWAIT := 5,
	ETT_WAITCINHRELEASE := 6,
	ETT_WAITCINH := 7,
	ETT_IDENTIFYTORQUE := 8,
	ETT_DONE := 10
);
END_TYPE

(* ---- L_MC1P_TOUCHPROBEINPUT.dut ---- *)
TYPE L_MC1P_TOUCHPROBEINPUT :
STRUCT
	EXECUTE : BOOL;
	WINDOWONLY : BOOL;
	FIRSTPOSITION : LREAL;
	LASTPOSITION : LREAL;
	PAUSEACTIVETP : BOOL;
	XBPB_S131_COMBINATION : BOOL;
END_STRUCT
END_TYPE

(* ---- L_MC1P_TOUCHPROBEOUTPUT.dut ---- *)
TYPE L_MC1P_TOUCHPROBEOUTPUT :
STRUCT
	DONE : BOOL;
	BUSY : BOOL;
	COMMANDABORTED : BOOL;
	ERROR : BOOL;
	ERRORID : L_IE1P_Error;
	ACTIVATIONLEVEL : BOOL;
	ACTIVATIONLEVELVALID : BOOL;
	VALUESTORED_POSEDGE : BOOL;
	RECPOSITION_POSEDGE : LREAL;
	VALUESTORED_NEGEDGE : BOOL;
	RECPOSITION_NEGEDGE : LREAL;
	NEWVALUESTORED_POSEDGE : BOOL;
	NEWVALUESTORED_NEGEDGE : BOOL;
	RECDATA : L_MC1P_TpReceiveData;
	TIMESTAMPFROMABSCOUNTERITF : L_IOM_IExternalTPInterface;
	TIMESTAMPABSCOUNTERHELPER : WORD;
END_STRUCT
END_TYPE

(* ---- L_MC1P_TPDATA.dut ---- *)
TYPE L_MC1P_TPDATA :
STRUCT
	XSTARTCAPTURING : BOOL;
	XINEXCECUTION : BOOL;
	XNEWEXECUTE : BOOL;
	XCOMMANDABORTED : BOOL;
	NERRORID : INT := 0;
	XVALUESTORED_POSEDGE : BOOL;
	DNRECORDEDPOSITION_POSEDGE : DINT;
	DWTIMESTAMP_POSEDGE : DWORD;
	XNEWVALUESTORED_POSEDGE : BOOL;
	XVALUESTORED_NEGEDGE : BOOL;
	DNRECORDEDPOSITION_NEGEDGE : DINT;
	DWTIMESTAMP_NEGEDGE : DWORD;
	XNEWVALUESTORED_NEGEDGE : BOOL;
	XACTIVATIONLEVEL : BOOL;
	XOVERRIDEACTIVE : BOOL;
	XTIMESTAMPAVAILABLEPOSEDGE : BOOL;
	XTIMESTAMPAVAILABLENEGEDGE : BOOL;
	XPOSITIONAVAILABLEPOSEDGE : BOOL;
	XPOSITIONAVAILABLENEGEDGE : BOOL;
	XACTIVATIONLEVELVALID : BOOL;
END_STRUCT
END_TYPE

(* ---- L_MC1P_TPRECEIVEDATA.dut ---- *)
TYPE L_MC1P_TPRECEIVEDATA :
STRUCT
	XVALUESTORED : BOOL;
	LRRECPOSITION : LREAL;
	DWRECTIMESTAMP : DWORD;
	DWACTTIMESTAMP : DWORD;
	XSUPPORTTIMESTAMP : BOOL;
	XSUPPORTPOSITION : BOOL;
	ITFTOUCHPROBEHANDLER : L_MC1P_ITouchProbeHandler;
	DWUPDATETIME : DWORD;
END_STRUCT
END_TYPE

(* ---- L_MC1P_TRAVERSINGRANGE.dut ---- *)
TYPE L_MC1P_TRAVERSINGRANGE :
(
	MODULO := 0,
	LIMITED := 1
);
END_TYPE

(* ---- L_MC1P_TRCELEMENT.dut ---- *)
TYPE L_MC1P_TRCELEMENT :
STRUCT
	DWCOUNT : DWORD;
	DWTRACEDATA_01 : DWORD;
	DWTRACEDATA_02 : DWORD;
	DWTRACEDATA_03 : DWORD;
	DWTRACEDATA_04 : DWORD;
	DWTRACEDATA_05 : DWORD;
	LRTRACEDATA_06 : LREAL;
	LRTRACEDATA_07 : LREAL;
	LRTRACEDATA_08 : LREAL;
END_STRUCT
END_TYPE

(* ---- L_MC1P_TYPEFUNCTION.dut ---- *)
TYPE L_MC1P_TYPEFUNCTION :
(
	TYPE_ANY := 0,
	TYPE_MC_MOVEABSOLUTE := 10,
	TYPE_MC_MOVEADDITIVE := 20,
	TYPE_MC_MOVECONTINUOUSABSOLUTE := 30,
	TYPE_MC_MOVECONTINUOUSRELATIVE := 40,
	TYPE_MC_MOVERELATIVE := 50,
	TYPE_MC_MOVESUPERIMPOSED := 60,
	TYPE_MC_HALTSUPERIMPOSED := 61,
	TYPE_MC_MOVEVELOCITY := 70,
	TYPE_MC_HALT := 80,
	TYPE_MC_STOP := 90,
	TYPE_MC_CAMIN := 100,
	TYPE_MC_CAMOUT := 110,
	TYPE_MC_GEARIN := 120,
	TYPE_MC_GEARINPOS := 130,
	TYPE_MC_GEAROUT := 140,
	TYPE_MC_COMBINEAXES := 150,
	TYPE_MC_PHASINGRELATIVE := 160,
	TYPE_MC_PHASINGABSOLUTE := 170,
	TYPE_MC_HOME := 180,
	TYPE_MC1P_FOLLOWSETVALUES := 190,
	TYPE_MC1P_TORQUECONTROL := 200,
	TYPE_CT1P_AUTOTUNING := 210,
	TYPE_MC1P_KINEMATICSYNC := 220
);
END_TYPE

(* ---- L_MC1P_UAXISRETAININFO.dut ---- *)
TYPE L_MC1P_UAXISRETAININFO :
UNION
	INFO : L_MC1P_AxisRetainInfo;
	DWDATA : DWORD;
END_UNION
END_TYPE

(* ---- L_MC1P_UNIVERSALAXISDATATYPES.dut ---- *)
TYPE L_MC1P_UNIVERSALAXISDATATYPES :
UNION
	AXISEXTENSION_I500_CAN : L_MC1P_AxisExtension_i500_CAN;
	AXISEXTENSION_I500_ECAT : L_MC1P_AxisExtension_i500_ECAT;
	AXISEXTENSION_I700 : L_MC1P_AxisExtension_i700;
	AXISEXTENSION_9400HL : L_MC1P_AxisExtension_9400HL;
	AXISEXTENSION_I750 : L_MC1P_AxisExtension_i750;
	AXISEXTENSION_I950 : L_MC1P_AxisExtension_i950;
	AXISEXTENSION_I950_CIAADV : L_MC1P_AxisExtension_i950_CiaAdv;
	AXISEXTENSION_GENERICDRIVE : L_MC1P_AxisExtension_GenericDrive;
END_UNION
END_TYPE

(* ---- L_MC1P_UNIVERSALENCODERDATATYPES.dut ---- *)
TYPE L_MC1P_UNIVERSALENCODERDATATYPES :
UNION
	AXISEXTENSION_ENCFREE : L_MC1P_AxisExtension_EncFree;
	AXISEXTENSION_ENCBPB : L_MC1P_AxisExtension_EncBPB;
	AXISEXTENSION_ENCI500 : L_MC1P_AxisExtension_Enci500;
	AXISEXTENSION_ENCI900_ECAT : L_MC1P_AxisExtension_Enci900_ECAT;
	AXISEXTENSION_ENCIOETC : L_MC1P_AxisExtension_EncIOEtc;
END_UNION
END_TYPE

(* ---- L_MC1P_UNSTEADYREASON.dut ---- *)
TYPE L_MC1P_UNSTEADYREASON :
(
	USRVIRTUAL := 0,
	USRREAL := 1,
	USRUNDEF := 9
);
END_TYPE

(* ---- L_MC1P_URETAINDATA.dut ---- *)
TYPE L_MC1P_URETAINDATA :
UNION
	RETAINDATAREALDRIVE : L_MC1P_RetainDataRealDrive_V3;
	RETAINDATAI700 : L_MC1P_RetainDatai700_V3;
END_UNION
END_TYPE

(* ---- L_MC1P_UULINT.dut ---- *)
TYPE L_MC1P_UULINT :
UNION
	ULIDATA : ULINT;
	AUDIDATA : ARRAY [1..2] OF UDINT;
END_UNION
END_TYPE

(* ---- L_MC1P_WRITEBOOLPARAMETERINPUT.dut ---- *)
TYPE L_MC1P_WRITEBOOLPARAMETERINPUT :
STRUCT
	EXECUTE : BOOL;
	PARAMETERNUMBER : DINT;
	VALUE : BOOL;
	EXECUTIONMODE : MC_EXECUTION_MODE;
END_STRUCT
END_TYPE

(* ---- L_MC1P_WRITEBOOLPARAMETEROUTPUT.dut ---- *)
TYPE L_MC1P_WRITEBOOLPARAMETEROUTPUT :
STRUCT
	DONE : BOOL;
	BUSY : BOOL;
	ERROR : BOOL;
	ERRORID : L_IE1P_Error;
END_STRUCT
END_TYPE

(* ---- L_MC1P_WRITEPARAMETERINPUT.dut ---- *)
TYPE L_MC1P_WRITEPARAMETERINPUT :
STRUCT
	AXIS : L_MC1P_IMCParameterAccess;
	EXECUTE : BOOL;
	PARAMETERNUMBER : DINT;
	VALUE : LREAL;
	EXECUTIONMODE : MC_EXECUTION_MODE;
END_STRUCT
END_TYPE

(* ---- L_MC1P_CONSTANTS.gvl ---- *)
VAR_GLOBAL
	GC_EPS : LREAL := 1E-10;
	GC_EPS_REAL : LREAL := 1E-06;
	GC_WUPDATEFILTER : WORD := 10;
	GC_WINSTANCENCHAR : WORD := 100;
	GC_WTRACEMAX : WORD := 100;
	GC_IMPLIZITCALLS : INT := 100;
	GC_MAXRETAINAXIS : INT := 256;
	GC_MAXAXISCOUNT : INT := 256;
	GC_ENCFILTERCYCLESMAX : INT := 100;
	GC_DWCHECKIDTAPPETREF : DWORD := 16#DC34;
	GC_SQRT2 : LREAL := 1.4142135623730951;
	GC_PI : LREAL := 3.1415926535897931;
	GC_REC_STATE : LWORD := SHL(1, 0);
	GC_REC_OPMODE : LWORD := SHL(1, 1);
	GC_REC_POS : LWORD := SHL(1, 2);
	GC_REC_VEL : LWORD := SHL(1, 3);
	GC_REC_TORQUE : LWORD := SHL(1, 4);
	GC_REC_ERRORID : LWORD := SHL(1, 5);
	GC_REC_FOLLERROR : LWORD := SHL(1, 6);
	GC_REC_STATELENZE : LWORD := SHL(1, 7);
	GC_REC_STATELENZE2 : LWORD := SHL(1, 8);
	GC_REC_TPSTATE1 : LWORD := SHL(1, 9);
	GC_REC_TP1POS : LWORD := SHL(1, 10);
	GC_REC_TP1NEG : LWORD := SHL(1, 11);
	GC_REC_TP2POS : LWORD := SHL(1, 12);
	GC_REC_TP2NEG : LWORD := SHL(1, 13);
	GC_REC_DIGIN : LWORD := SHL(1, 14);
	GC_REC_STATESM : LWORD := SHL(1, 15);
	GC_REC_VLACTVELOCITY : LWORD := SHL(1, 16);
	GC_REC_ENCPOS : LWORD := SHL(1, 17);
	GC_REC_ENCVEL : LWORD := SHL(1, 18);
	GC_REC_TP1POSTIME : LWORD := SHL(1, 19);
	GC_REC_TP1NEGTIME : LWORD := SHL(1, 20);
	GC_REC_TP2POSTIME : LWORD := SHL(1, 21);
	GC_REC_TP2NEGTIME : LWORD := SHL(1, 22);
	GC_REC_TPSTATE2 : LWORD := SHL(1, 23);
	GC_REC_TP3POS : LWORD := SHL(1, 24);
	GC_REC_TP3NEG : LWORD := SHL(1, 25);
	GC_REC_TP4POS : LWORD := SHL(1, 26);
	GC_REC_TP4NEG : LWORD := SHL(1, 27);
	GC_REC_TP3POSTIME : LWORD := SHL(1, 28);
	GC_REC_TP3NEGTIME : LWORD := SHL(1, 29);
	GC_REC_TP4POSTIME : LWORD := SHL(1, 30);
	GC_REC_TP4NEGTIME : LWORD := SHL(1, 31);
	GC_REC_SAFETYCTRL : LWORD := SHL(1, 32);
	GC_REC_SAFETYSTATE : LWORD := SHL(1, 33);
	GC_REC_SAFETYIOSTATE : LWORD := SHL(1, 34);
	GC_REC_ENCPOSTIMESTAMP : LWORD := SHL(1, 35);
	GC_REC_STATELENZEEXT : LWORD := SHL(1, 36);
	GC_REC_SPEEDERROR : LWORD := SHL(1, 37);
	GC_REC_POSVALUE1616 : LWORD := SHL(1, 38);
	GC_REC_CONTROLEFFORT : LWORD := SHL(1, 39);
	GC_REC_ACTPOSMOTORCIA402ADV : LWORD := SHL(1, 40);
	GC_REC_TEXTREFID : LWORD := SHL(1, 41);
	GC_REC_POSTIMESTAMP : LWORD := SHL(1, 42);
	GC_REC_MAXDATAINDEX : WORD := 43;
	GC_TRANS_CTRL : LWORD := SHL(1, 0);
	GC_TRANS_OPMODE : LWORD := SHL(1, 1);
	GC_TRANS_POS : LWORD := SHL(1, 2);
	GC_TRANS_VEL : LWORD := SHL(1, 3);
	GC_TRANS_TORQUE : LWORD := SHL(1, 4);
	GC_TRANS_TORQUELIMPOS : LWORD := SHL(1, 5);
	GC_TRANS_TORQUELIMNEG : LWORD := SHL(1, 6);
	GC_TRANS_SPEEDLIMUP : LWORD := SHL(1, 7);
	GC_TRANS_SPEEDLIMLOW : LWORD := SHL(1, 8);
	GC_TRANS_TPCTRL1 : LWORD := SHL(1, 9);
	GC_TRANS_POSOFFSET : LWORD := SHL(1, 10);
	GC_TRANS_VELOFFSET : LWORD := SHL(1, 11);
	GC_TRANS_TORQUEOFFSET : LWORD := SHL(1, 12);
	GC_TRANS_SPEEDCTRLINT : LWORD := SHL(1, 13);
	GC_TRANS_CTRLLENZE : LWORD := SHL(1, 14);
	GC_TRANS_VLTARGETVELOCITY : LWORD := SHL(1, 16);
	GC_TRANS_BRKOVRD : LWORD := SHL(1, 17);
	GC_TRANS_CTRLLENZE2 : LWORD := SHL(1, 18);
	GC_TRANS_CTRLLENZE3 : LWORD := SHL(1, 19);
	GC_TRANS_CTRLLENZE4 : LWORD := SHL(1, 20);
	GC_TRANS_TPCTRL2 : LWORD := SHL(1, 21);
	GC_TRANS_SAFEPOS : LWORD := SHL(1, 22);
	GC_TRANS_SAFEPOSSTATUS : LWORD := SHL(1, 23);
	GC_TRANS_SPEEDLIMITSLS : LWORD := SHL(1, 24);
	GC_TRANS_MAXDATAINDEX : WORD := 25;
	NODATAMEMORYAVAILABLE : WORD := WORD#16#1;
	MEMORYINVALID : WORD := WORD#16#2;
	MEMORYNOTINITIALIZED : WORD := WORD#16#4;
	NODATAAVAILABLE : WORD := WORD#16#8;
	NOMEMORYAVAILABLEFORAXIS : WORD := WORD#16#10;
	NOMEMORYINAXISARRAY : WORD := WORD#16#20;
	AXISGUIDCHANGED : WORD := WORD#16#40;
	C_SERIALNUMBER : UINT := 3;
	C_MANUFACTURER : UINT := 5;
	C_SOFTWAREREVISION : UINT := 9;
	C_HARDWAREREVISION : UINT := 10;
	C_DEVICECLASS : UINT := 11;
	C_PRODUCTCODE : UINT := 13;
	C_UPDATE : UINT := 99;
	C_CONNECTORTYPEMOTIONAXISOLD : UINT := 1279;
	C_CONNECTORTYPEMOTIONAXIS : UINT := 34279;
	C_CONNECTORTYPEENCODERIOSLICE : UINT := 33024;
END_VAR

(* ---- L_MC1P_INTERNAL.gvl ---- *)
VAR_GLOBAL
	DWDUMMY : DWORD;
	XAPPFIRSTRUN : BOOL := FALSE;
	PANYCONNECTOR : POINTER TO IoConfigConnector;
	LMAXISRETAINHANDLING : L_MC1P_AxisRetainMangaement;
	DWTIMESTAMPSIMU : DWORD;
	XTIMESTAMPUPDATED : BOOL;
	LMAXISMGMT : L_MC1P_AxisManagementFunction;
	CDIENUMSTARTVALUE : DINT := 50000;
END_VAR

(* ---- L_MC1P_IAXIS_REF_BRAKE.itf ---- *)
INTERFACE L_MC1P_IAXIS_REF_BRAKE
END_INTERFACE

METHOD GETACTVALUESBRAKE
END_METHOD

METHOD SWITCHONCONTROL
VAR_INPUT
	XSWITCHONREQUEST : BOOL;
END_VAR
VAR_OUTPUT
	XSWITCHON : BOOL;
END_VAR
VAR_IN_OUT
	AXIS : AXIS_REF;
END_VAR
END_METHOD

METHOD SWITCHEDONSTATUS
VAR_INPUT
	XSWITCHEDONREQUEST : BOOL;
END_VAR
VAR_OUTPUT
	XSWITCHEDON : BOOL;
END_VAR
VAR_IN_OUT
	AXIS : AXIS_REF;
END_VAR
END_METHOD

(* ---- L_MC1P_IAXIS_REF_MASTERVALUES.itf ---- *)
INTERFACE L_MC1P_IAXIS_REF_MASTERVALUES
END_INTERFACE

METHOD GETDIRECTION : WORD
VAR_INPUT
	VALUESOURCE : MC_SOURCE;
END_VAR
END_METHOD

METHOD GETMASTERERROR : BOOL
VAR_OUTPUT
	EERRORID : L_IE1P_Error;
END_VAR
END_METHOD

METHOD GETSTEADYSTATE : POINTER TO L_MC1P_SteadyState
END_METHOD

(* ---- L_MC1P_IAXIS_REF_POOL.itf ---- *)
INTERFACE L_MC1P_IAXIS_REF_POOL
END_INTERFACE

METHOD GETAXISFROMPOOL : POINTER TO AXIS_REF
VAR_INPUT
	WINDEX : WORD;
END_VAR
END_METHOD
